// ---- 10_Core/90_Redundancy/FB_RedSync.TcPOU
FUNCTION_BLOCK FB_RedSync		// 동기화: 이 PLC의 운영 설정(GVL_PERSIST, 모듈 설정 묶음 제외)과 제어 모드 요청(PCS마다)을 EAP로 매 스캔 상대에게 보내고, 상대가 Active이고 내가 Active가 아닐 때 받은 값으로 내 설정을 맞춘다
(* - 보내는 값은 EAP 변수 1개: 운영 설정(_stTx, ST_RedSyncCfg). 받는 값도 같은 모양(_stRx)
   - 모듈 설정 묶음(GVL_PERSIST.g_stModuleSet)은 동기화하지 않음: HMI가 두 PLC 모두에 씀 (PLC가 꺼져 있던 동안 바꾼 값은 복귀 전에 HMI에서 다시 쓸 것)
   - 맞추기: i_bApply일 때만, 값이 다른 것만 덮어씀 (같으면 안 씀: 저장을 불필요하게 만들지 않음). 바꾼 것이 없으면 q_bInSync
   - 살아 있음: _stRx.nSeq가 i_tTimeout 안에 바뀌어야 함 (q_bFresh)
   - I/O(AT %I*·%Q)는 설치할 때 XAE에서 연결. 인스턴스는 RedundancyTask의 PRG_Redundancy에 둠. 두 PLC 프로그램이 같아야 함 *)
VAR_INPUT
	i_bUse			: BOOL;
	i_bApply		: BOOL;				// 받은 값을 내 설정에 덮어써도 됨 (내가 Active가 아니고 상대가 Active이며 통신 정상)
	i_tTimeout		: TIME := T#2S;		// 새 값이 이 시간 안에 안 오면 낡은 것
END_VAR
VAR_OUTPUT
	q_bInSync		: BOOL;				// 받은 값이 낡지 않았고 내 설정이 그와 같음 (i_bApply일 때만 TRUE)
	q_bFresh		: BOOL;				// 상대가 보낸 값이 낡지 않음
	q_nApplied		: UDINT;			// 받은 값으로 덮어쓴 횟수 (필드 단위)
END_VAR
VAR
	(* I/O: XAE에서 연결 *)
	_stTx			AT %Q* : ST_RedSyncCfg;
	_stRx			AT %I* : ST_RedSyncCfg;

	_nLastSeq		: UDINT;
	_tonFresh		: TON;
END_VAR
VAR_TEMP
	bNew			: BOOL;
	bEq				: BOOL;
END_VAR

IF NOT i_bUse THEN
	RETURN;
END_IF

(* 1) 보내기 *)
_stTx.nProtoVer	:= 1;
_stTx.nSeq		:= _stTx.nSeq + 1;
_stTx.nModeReq1	:= GVL_SITE.g_fbCtrlMode1.i_nModeReq;
_stTx.aeOpMode := GVL_PERSIST.g_aeOpMode;
_stTx.astGroupSet := GVL_PERSIST.g_astGroupSet;
_stTx.astManualPolicy := GVL_PERSIST.g_astManualPolicy;
_stTx.astSourceReg := GVL_PERSIST.g_astSourceReg;
_stTx.astLimitReg := GVL_PERSIST.g_astLimitReg;
_stTx.astPermitReg := GVL_PERSIST.g_astPermitReg;
_stTx.astCompReg := GVL_PERSIST.g_astCompReg;
_stTx.astRuleCfg := GVL_PERSIST.g_astRuleCfg;
_stTx.astOutputCfg := GVL_PERSIST.g_astOutputCfg;
_stTx.astUnitRuleReg := GVL_PERSIST.g_astUnitRuleReg;
_stTx.astBatRuleReg := GVL_PERSIST.g_astBatRuleReg;
_stTx.stCmdFilter := GVL_PERSIST.g_stCmdFilter;
_stTx.stManualCmdSet := GVL_PERSIST.g_stManualCmdSet;
_stTx.stSeqSet := GVL_PERSIST.g_stSeqSet;
_stTx.stBrokerWatch := GVL_PERSIST.g_stBrokerWatch;	// [9번 수정 2026-11-09: 추가]

(* 2) 받기: 새 값이 오는지 *)
bNew := _stRx.nSeq <> _nLastSeq;
_nLastSeq := _stRx.nSeq;
_tonFresh(IN := NOT bNew, PT := i_tTimeout);
q_bFresh := _stRx.nProtoVer = 1 AND _stRx.nSeq <> 0 AND NOT _tonFresh.Q;

(* 3) 맞추기: 내가 Active가 아니고 상대가 Active일 때만 다른 것만 덮어씀 *)
q_bInSync := FALSE;
IF i_bApply AND q_bFresh THEN
	bEq := TRUE;
	IF GVL_SITE.g_fbCtrlMode1.i_nModeReq <> _stRx.nModeReq1 THEN
		GVL_SITE.g_fbCtrlMode1.i_nModeReq := _stRx.nModeReq1;
		q_nApplied := q_nApplied + 1;
		bEq := FALSE;
	END_IF
	IF MEMCMP(ADR(GVL_PERSIST.g_aeOpMode), ADR(_stRx.aeOpMode), SIZEOF(_stRx.aeOpMode)) <> 0 THEN
		GVL_PERSIST.g_aeOpMode := _stRx.aeOpMode;
		q_nApplied := q_nApplied + 1;
		bEq := FALSE;
	END_IF
	IF MEMCMP(ADR(GVL_PERSIST.g_astGroupSet), ADR(_stRx.astGroupSet), SIZEOF(_stRx.astGroupSet)) <> 0 THEN
		GVL_PERSIST.g_astGroupSet := _stRx.astGroupSet;
		q_nApplied := q_nApplied + 1;
		bEq := FALSE;
	END_IF
	IF MEMCMP(ADR(GVL_PERSIST.g_astManualPolicy), ADR(_stRx.astManualPolicy), SIZEOF(_stRx.astManualPolicy)) <> 0 THEN
		GVL_PERSIST.g_astManualPolicy := _stRx.astManualPolicy;
		q_nApplied := q_nApplied + 1;
		bEq := FALSE;
	END_IF
	IF MEMCMP(ADR(GVL_PERSIST.g_astSourceReg), ADR(_stRx.astSourceReg), SIZEOF(_stRx.astSourceReg)) <> 0 THEN
		GVL_PERSIST.g_astSourceReg := _stRx.astSourceReg;
		q_nApplied := q_nApplied + 1;
		bEq := FALSE;
	END_IF
	IF MEMCMP(ADR(GVL_PERSIST.g_astLimitReg), ADR(_stRx.astLimitReg), SIZEOF(_stRx.astLimitReg)) <> 0 THEN
		GVL_PERSIST.g_astLimitReg := _stRx.astLimitReg;
		q_nApplied := q_nApplied + 1;
		bEq := FALSE;
	END_IF
	IF MEMCMP(ADR(GVL_PERSIST.g_astPermitReg), ADR(_stRx.astPermitReg), SIZEOF(_stRx.astPermitReg)) <> 0 THEN
		GVL_PERSIST.g_astPermitReg := _stRx.astPermitReg;
		q_nApplied := q_nApplied + 1;
		bEq := FALSE;
	END_IF
	IF MEMCMP(ADR(GVL_PERSIST.g_astCompReg), ADR(_stRx.astCompReg), SIZEOF(_stRx.astCompReg)) <> 0 THEN
		GVL_PERSIST.g_astCompReg := _stRx.astCompReg;
		q_nApplied := q_nApplied + 1;
		bEq := FALSE;
	END_IF
	IF MEMCMP(ADR(GVL_PERSIST.g_astRuleCfg), ADR(_stRx.astRuleCfg), SIZEOF(_stRx.astRuleCfg)) <> 0 THEN
		GVL_PERSIST.g_astRuleCfg := _stRx.astRuleCfg;
		q_nApplied := q_nApplied + 1;
		bEq := FALSE;
	END_IF
	IF MEMCMP(ADR(GVL_PERSIST.g_astOutputCfg), ADR(_stRx.astOutputCfg), SIZEOF(_stRx.astOutputCfg)) <> 0 THEN
		GVL_PERSIST.g_astOutputCfg := _stRx.astOutputCfg;
		q_nApplied := q_nApplied + 1;
		bEq := FALSE;
	END_IF
	IF MEMCMP(ADR(GVL_PERSIST.g_astUnitRuleReg), ADR(_stRx.astUnitRuleReg), SIZEOF(_stRx.astUnitRuleReg)) <> 0 THEN
		GVL_PERSIST.g_astUnitRuleReg := _stRx.astUnitRuleReg;
		q_nApplied := q_nApplied + 1;
		bEq := FALSE;
	END_IF
	IF MEMCMP(ADR(GVL_PERSIST.g_astBatRuleReg), ADR(_stRx.astBatRuleReg), SIZEOF(_stRx.astBatRuleReg)) <> 0 THEN
		GVL_PERSIST.g_astBatRuleReg := _stRx.astBatRuleReg;
		q_nApplied := q_nApplied + 1;
		bEq := FALSE;
	END_IF
	IF MEMCMP(ADR(GVL_PERSIST.g_stCmdFilter), ADR(_stRx.stCmdFilter), SIZEOF(_stRx.stCmdFilter)) <> 0 THEN
		GVL_PERSIST.g_stCmdFilter := _stRx.stCmdFilter;
		q_nApplied := q_nApplied + 1;
		bEq := FALSE;
	END_IF
	IF MEMCMP(ADR(GVL_PERSIST.g_stManualCmdSet), ADR(_stRx.stManualCmdSet), SIZEOF(_stRx.stManualCmdSet)) <> 0 THEN
		GVL_PERSIST.g_stManualCmdSet := _stRx.stManualCmdSet;
		q_nApplied := q_nApplied + 1;
		bEq := FALSE;
	END_IF
	IF MEMCMP(ADR(GVL_PERSIST.g_stSeqSet), ADR(_stRx.stSeqSet), SIZEOF(_stRx.stSeqSet)) <> 0 THEN
		GVL_PERSIST.g_stSeqSet := _stRx.stSeqSet;
		q_nApplied := q_nApplied + 1;
		bEq := FALSE;
	END_IF
	IF MEMCMP(ADR(GVL_PERSIST.g_stBrokerWatch), ADR(_stRx.stBrokerWatch), SIZEOF(_stRx.stBrokerWatch)) <> 0 THEN	// [9번 수정 2026-11-09: 추가]
		GVL_PERSIST.g_stBrokerWatch := _stRx.stBrokerWatch;
		q_nApplied := q_nApplied + 1;
		bEq := FALSE;
	END_IF
	q_bInSync := bEq;
END_IF

END_FUNCTION_BLOCK

// ---- 10_Core/90_Redundancy/FB_RedState.TcPOU
FUNCTION_BLOCK FB_RedState		// 이중화 상태 기계 (순수 로직). 역할 + 상대 상태 → 이 PLC가 Active인지, 장비에 써도 되는지. 두 PLC가 동시에 Active가 되지 않게 함
(* 규칙
   - 이중화를 안 쓰면 항상 Active이고 바로 쓴다
   - 역할 설정 오류(NoMatch) 또는 두 PLC 역할이 같음 → Failed (둘 다 장비에 쓰지 않음)
   - Primary: 시작하면 상대 상태를 볼 때까지 Init. 상대가 Active가 아니면 Active, 이미 Active이면 뺏지 않고 Standby
   - 절체: Secondary는 상대가 Lost(EAP·접점 둘 다 끊김)이고 tTakeoverDelay가 지나면 Active (Standby → Active)
   - 복귀: Primary가 Standby에서 상대(Secondary)가 Active이고 통신이 tFailbackStable 동안 정상이면 Handover(넘겨받기 요청)로 감.
     Secondary는 상대가 Handover이면 Active를 내려놓고 Standby로. Primary는 상대가 Active가 아니게 되면 Active.
     tHandoverTimeout 안에 안 내려놓으면 Primary가 Standby로 돌아가 다시 기다림. 둘 다 안 쓰는 틈이 생기지만 둘 다 쓰는 일은 없음
   - 둘 다 Active로 보이면 Secondary가 Standby로 물러남 (Primary 우선)
   - 상대 Active = EAP 하트비트의 Active (EAP 정상일 때) 또는 Active 접점 (접점 정상일 때)
   - PLC가 멈췄다 이어지면(i_bReset) Init부터 다시 정함: 멈춘 사이 상대가 Active를 넘겨받았을 수 있으므로 옛 Active를 이어 쓰지 않고, 상대 상태를 본 뒤 Standby로 들어가 복귀 절차를 밟음
   - 장비에 쓰는 허가(q_bWrite)는 Active가 된 뒤 tWriteHold가 지나야 켜짐 (승격 직후 계산이 안정되기를 기다림). Active가 아니게 되면 바로 꺼짐 *)
VAR_INPUT
	i_bUse			: BOOL;				// GVL_SITE.RED_SET.bUse
	i_stSet			: ST_RedSet;		// 시간 설정
	i_eRole			: E_RedRole;
	i_ePeer			: E_RedPeer;
	i_bPeerActive	: BOOL;				// 상대가 Active (EAP 또는 접점. 정상인 쪽만 반영해서 넘길 것)
	i_bPeerHandover	: BOOL;				// 상대가 Handover라고 알림 (EAP 정상일 때만)
	i_bRoleConflict	: BOOL;				// 두 PLC 역할이 같음 (FB_RedPeerMonitor)
	i_bReset		: BOOL;				// PLC가 멈췄다 이어짐: 상태를 Init부터 다시 정함 (멈춘 사이 상대가 Active를 넘겨받았을 수 있음)
	i_bSyncDone		: BOOL := TRUE;		// 복귀 전에 상대에게서 받을 값 동기화가 끝났음 (4단계에서 연결. 지금은 항상 TRUE)
END_VAR
VAR_OUTPUT
	q_eState		: E_RedState;
	q_bActive		: BOOL;				// Active 상태 (상대에게 알림)
	q_bWrite		: BOOL;				// 장비에 써도 됨 (Active + 쓰기 대기 지남)
	q_nSwitchCount	: UDINT;			// Active가 바뀐 횟수 (들어가거나 나옴)
	q_eLastSwitch	: E_RedSwitch;		// 마지막으로 바뀐 이유
END_VAR
VAR
	_ePrev			: E_RedState;
	_tonTakeover	: TON;
	_tonFailback	: TON;
	_tonHandover	: TON;
	_tonHold		: TON;
END_VAR

// 타이머는 매 스캔 부름
_tonTakeover(IN := i_eRole = E_RedRole.Secondary AND q_eState = E_RedState.Standby AND i_ePeer = E_RedPeer.Lost, PT := i_stSet.tTakeoverDelay);
_tonFailback(IN := i_eRole = E_RedRole.Primary AND q_eState = E_RedState.Standby AND i_ePeer = E_RedPeer.Alive AND i_bPeerActive AND i_bSyncDone, PT := i_stSet.tFailbackStable);
_tonHandover(IN := q_eState = E_RedState.Handover, PT := i_stSet.tHandoverTimeout);

IF i_bReset THEN
	q_eState := E_RedState.Init;
ELSIF NOT i_bUse THEN
	q_eState := E_RedState.Active;
ELSIF i_eRole = E_RedRole.NoMatch OR i_bRoleConflict THEN
	q_eState := E_RedState.Failed;
ELSIF i_eRole = E_RedRole.Reading THEN
	q_eState := E_RedState.Init;
ELSE
	IF q_eState = E_RedState.Failed THEN
		q_eState := E_RedState.Init;		// 오류가 풀리면 처음부터 다시 정함
	END_IF
	CASE q_eState OF
	E_RedState.Init:
		IF i_eRole = E_RedRole.Secondary THEN
			q_eState := E_RedState.Standby;
		ELSIF i_ePeer <> E_RedPeer.Unknown THEN		// Primary: 상대 상태를 본 뒤 정함
			IF i_bPeerActive THEN
				q_eState := E_RedState.Standby;
			ELSE
				q_eState := E_RedState.Active;
				q_eLastSwitch := E_RedSwitch.Start;
			END_IF
		END_IF
	E_RedState.Standby:
		IF i_eRole = E_RedRole.Secondary THEN
			IF _tonTakeover.Q THEN
				q_eState := E_RedState.Active;		// 절체
				q_eLastSwitch := E_RedSwitch.PeerLost;
			END_IF
		ELSIF i_ePeer <> E_RedPeer.Unknown THEN		// Primary
			IF NOT i_bPeerActive THEN
				q_eState := E_RedState.Active;		// 상대가 Active가 아님 (정지·대기)
				q_eLastSwitch := E_RedSwitch.Start;
			ELSIF _tonFailback.Q THEN
				q_eState := E_RedState.Handover;	// 복귀: 상대에게 Active를 내려놓으라고 알림
			END_IF
		END_IF
	E_RedState.Handover:
		IF NOT i_bPeerActive THEN
			q_eState := E_RedState.Active;			// 상대가 내려놓음 (또는 사라짐)
			q_eLastSwitch := E_RedSwitch.Failback;
		ELSIF _tonHandover.Q OR i_ePeer <> E_RedPeer.Alive THEN
			q_eState := E_RedState.Standby;			// 포기하고 처음부터 다시 기다림
		END_IF
	E_RedState.Active:
		IF i_eRole = E_RedRole.Secondary AND (i_bPeerActive OR i_bPeerHandover) THEN
			q_eState := E_RedState.Standby;			// Primary에 양보
			q_eLastSwitch := E_RedSwitch.Yield;
		END_IF
	ELSE
		q_eState := E_RedState.Init;
	END_CASE
END_IF

// Active가 들어가거나 나올 때 횟수
IF (q_eState = E_RedState.Active) <> (_ePrev = E_RedState.Active) THEN
	q_nSwitchCount := q_nSwitchCount + 1;
END_IF
_ePrev := q_eState;

q_bActive := q_eState = E_RedState.Active;
_tonHold(IN := q_bActive, PT := i_stSet.tWriteHold);
q_bWrite := q_bActive AND (_tonHold.Q OR NOT i_bUse);

END_FUNCTION_BLOCK

// ---- 10_Core/90_Redundancy/FB_RedLink.TcPOU
FUNCTION_BLOCK FB_RedLink		// 이중화 연결: EAP 하트비트 보내기·받기 + 접점 신호(EL2004 출력·EL1004 입력) 보내기·받기 + 상대 상태 판정 (FB_RedPeerMonitor)
(* - I/O 연결(AT %I*·%Q)은 설치할 때 XAE에서 한다. 인스턴스는 RedundancyTask를 도는 PRG_Redundancy에 둔다
   - EAP 보내기 _stTx → 상대가 받음, 받기 _stRx ← 상대가 보냄, Quality _nEapQuality: EAP 변수 연결 (값 = 마지막 갱신 뒤 지난 시간, 100 us 단위)
   - 접점: _bDoAlive(EL2004 채널 1)는 주기적으로 뒤집음 → 상대 _bDiPeerAlive(EL1004 채널 1). _bDoActive(채널 2)는 이 PLC가 Active인 동안 TRUE → 상대 _bDiPeerActive(채널 2)
   - 두 PLC에 같은 프로그램을 넣고, 두 PLC의 I/O 연결이 서로 마주 보게 한다 *)
VAR_INPUT
	i_stSet			: ST_RedSet;
	i_eRole			: E_RedRole;
	i_bActive		: BOOL;
	i_eState		: E_RedState;		// 이 PLC의 이중화 상태 (상대에게 알림)
END_VAR
VAR_OUTPUT
	q_ePeer			: E_RedPeer;		// 상대 상태
	q_bEapOk		: BOOL;
	q_bWireOk		: BOOL;
	q_stPeer		: ST_RedHeartbeat;	// 상대가 보낸 역할·Active (EAP 정상일 때만)
	q_bPeerWireActive: BOOL;			// 상대 Active 접점 (EAP와 따로 보는 값)
	q_bRoleConflict	: BOOL;				// 두 PLC 역할이 같음
	q_nTxCount		: UDINT;			// 보낸 하트비트 수
END_VAR
VAR CONSTANT
	PULSE_HALF		: TIME := T#100MS;	// alive 접점을 뒤집는 간격 (접점 타임아웃보다 충분히 짧게)
END_VAR
VAR
	(* I/O: XAE에서 연결 *)
	_stTx			AT %Q* : ST_RedHeartbeat;
	_stRx			AT %I* : ST_RedHeartbeat;
	_nEapQuality	AT %I* : UINT;		// EAP Subscriber의 Quality = 갱신 안 된 시간 (100 us 단위). tEapTimeout 이하면 정상
	_bDoAlive		AT %Q* : BOOL;		// EL2004 채널 1
	_bDoActive		AT %Q* : BOOL;		// EL2004 채널 2
	_bDiPeerAlive	AT %I* : BOOL;		// EL1004 채널 1
	_bDiPeerActive	AT %I* : BOOL;		// EL1004 채널 2

	_fbMon			: FB_RedPeerMonitor;
	_tonPulse		: TON;
END_VAR

(* 1) 보내기 *)
q_nTxCount			:= q_nTxCount + 1;
_stTx.nProtoVer		:= 2;
_stTx.nCounter		:= q_nTxCount;
_stTx.nRole			:= TO_INT(i_eRole);
_stTx.bActive		:= i_bActive;
_stTx.nState		:= TO_INT(i_eState);

_tonPulse(IN := NOT _tonPulse.Q, PT := PULSE_HALF);		// Q가 한 스캔 켜질 때마다 뒤집음
IF _tonPulse.Q THEN
	_bDoAlive := NOT _bDoAlive;
END_IF
_bDoActive			:= i_bActive;

(* 2) 받아서 판정 *)
_fbMon(	i_stRx			:= _stRx,
		i_nMyRole		:= TO_INT(i_eRole),
		i_bEapQualityOk	:= UINT_TO_UDINT(_nEapQuality) <= TIME_TO_UDINT(i_stSet.tEapTimeout) * 10,	// Quality = 갱신 안 된 시간 (100 us 단위)
		i_bWireAlive	:= _bDiPeerAlive,
		i_tEapTimeout	:= i_stSet.tEapTimeout,
		i_tWireTimeout	:= i_stSet.tWireTimeout,
		i_tStartGrace	:= i_stSet.tStartGrace);
q_ePeer				:= _fbMon.q_ePeer;
q_bEapOk			:= _fbMon.q_bEapOk;
q_bWireOk			:= _fbMon.q_bWireOk;
q_stPeer			:= _fbMon.q_stPeer;
q_bPeerWireActive	:= _bDiPeerActive;
q_bRoleConflict		:= _fbMon.q_bRoleConflict;

END_FUNCTION_BLOCK

// ---- 10_Core/90_Redundancy/FB_RedPeerMonitor.TcPOU
FUNCTION_BLOCK FB_RedPeerMonitor		// 상대 PLC 상태 판정 (순수 로직: I/O를 직접 안 봄). EAP 하트비트(카운터가 바뀌고 Quality 정상)와 접점 신호(값이 바뀜)를 따로 보고 합침
// 판정 규칙: 둘 다 정상 = Alive, 한쪽만 끊김 = 그 통신 고장 (상대는 살아 있음, 절체 안 함), 둘 다 끊김 = Lost (절체 조건)
VAR_INPUT
	i_stRx			: ST_RedHeartbeat;	// 받은 EAP 하트비트
	i_bEapQualityOk	: BOOL;				// EAP Quality가 정상
	i_nMyRole		: INT;				// 이 PLC의 역할 (E_RedRole). 받은 역할이 같으면 내 프레임이 되돌아온 것으로 보고 무시
	i_bWireAlive	: BOOL;				// 상대 alive 접점(DI)의 지금 값. 상대가 주기적으로 뒤집음
	i_tEapTimeout	: TIME := T#500MS;	// 카운터가 이 시간 안 바뀌면 EAP 끊김
	i_tWireTimeout	: TIME := T#500MS;	// 접점이 이 시간 안 바뀌면 접점 끊김
	i_tStartGrace	: TIME := T#3S;		// 시작 직후 대기: 이 안에는 아직 못 봐도 Unknown
END_VAR
VAR_OUTPUT
	q_ePeer			: E_RedPeer;
	q_bEapOk		: BOOL;				// EAP 하트비트 정상
	q_bWireOk		: BOOL;				// 접점 신호 정상
	q_stPeer		: ST_RedHeartbeat;	// 상대가 보낸 값. EAP가 정상일 때만 채움 (아니면 0)
	q_bRoleConflict	: BOOL;				// 상대가 나와 같은 역할로 살아 있음 (두 PLC 역할 설정 오류). 접점도 살아 있을 때만 (내 프레임이 되돌아온 경우와 구분)
END_VAR
VAR
	_bInit			: BOOL;
	_nLastCount		: UDINT;
	_bLastWire		: BOOL;
	_bEapSeen		: BOOL;			// 시작 뒤 카운터가 바뀌는 것을 한 번이라도 봄
	_bWireSeen		: BOOL;
	_bSameSeen		: BOOL;
	_tonSame		: TON;
	_tonEap			: TON;
	_tonWire		: TON;
	_tonStart		: TON;
END_VAR
VAR_TEMP
	bEapMoved		: BOOL;
	bFromSelf		: BOOL;
	bSameMoved		: BOOL;
	bCntMoved		: BOOL;
	bWireMoved		: BOOL;
	stZero			: ST_RedHeartbeat;
END_VAR

IF NOT _bInit THEN
	_nLastCount	:= i_stRx.nCounter;
	_bLastWire	:= i_bWireAlive;
	_bInit		:= TRUE;
END_IF

// EAP: 카운터가 바뀌었고 Quality 정상이면 살아 있음. 안 바뀌는 시간이 길면 끊김 (상대 PLC가 멈추면 마지막 값이 그대로 남으므로 Quality만으로는 못 잡음)
bFromSelf		:= i_stRx.nRole = i_nMyRole;	// 상대와 내 역할은 항상 다름. 같으면 루프로 되돌아온 내 프레임 (또는 역할 설정 오류)
bCntMoved		:= i_bEapQualityOk AND i_stRx.nCounter <> _nLastCount;
bEapMoved		:= bCntMoved AND NOT bFromSelf;
_nLastCount		:= i_stRx.nCounter;
IF bEapMoved THEN
	_bEapSeen := TRUE;
END_IF
// 같은 역할 프레임이 계속 오는지 (Primary·Secondary일 때만. 시작 중 Reading끼리는 제외)
bSameMoved		:= bCntMoved AND bFromSelf AND (i_nMyRole = 1 OR i_nMyRole = 2);
IF bSameMoved THEN
	_bSameSeen := TRUE;
END_IF
_tonSame(IN := NOT bSameMoved, PT := i_tEapTimeout);
_tonEap(IN := NOT bEapMoved, PT := i_tEapTimeout);
q_bEapOk		:= _bEapSeen AND NOT _tonEap.Q AND i_bEapQualityOk AND NOT bFromSelf;

// 접점: 값이 바뀌면 살아 있음
bWireMoved		:= i_bWireAlive <> _bLastWire;
_bLastWire		:= i_bWireAlive;
IF bWireMoved THEN
	_bWireSeen := TRUE;
END_IF
_tonWire(IN := NOT bWireMoved, PT := i_tWireTimeout);
q_bWireOk		:= _bWireSeen AND NOT _tonWire.Q;
q_bRoleConflict	:= _bSameSeen AND NOT _tonSame.Q AND q_bWireOk;

_tonStart(IN := TRUE, PT := i_tStartGrace);

IF q_bEapOk AND q_bWireOk THEN
	q_ePeer := E_RedPeer.Alive;
ELSIF q_bWireOk THEN
	q_ePeer := E_RedPeer.EapLost;
ELSIF q_bEapOk THEN
	q_ePeer := E_RedPeer.WireLost;
ELSIF NOT _bEapSeen AND NOT _bWireSeen AND NOT _tonStart.Q THEN
	q_ePeer := E_RedPeer.Unknown;
ELSE
	q_ePeer := E_RedPeer.Lost;
END_IF

IF q_bEapOk THEN
	q_stPeer := i_stRx;
ELSE
	q_stPeer := stZero;
END_IF

END_FUNCTION_BLOCK

// ---- 20_Module/Common/FB_AuxIo.TcPOU
FUNCTION_BLOCK FB_AuxIo EXTENDS FB_DeviceBase IMPLEMENTS I_AuxDevice		// 벡호프 단자 I/O (EL1xxx 입력, EL2xxx 출력, EL3xxx 아날로그 입력, EL4xxx 아날로그 출력)
(* 점은 TwinCAT 화면에서 _abDi·_abDo·_anAi·_anAo 칸에 하나씩 연결. 점 번호 = 배열 칸 번호
   이 FB를 PlcTask가 아닌 태스크에서 쓰면 그 태스크 PRG 안에 선언 (GVL에 두면 TcContextName 필요) *)
VAR_INPUT
	i_afAiGain		: ARRAY[1..GVL_PARAM.AUX_AI_MAX] OF REAL;		// 아날로그 입력 = 원시값 × 배율 + 오프셋. 배율 0 = 1 (예: PT100 EL3202는 0.1)
	i_afAiOffset	: ARRAY[1..GVL_PARAM.AUX_AI_MAX] OF REAL;
	i_afAoGain		: ARRAY[1..GVL_PARAM.AUX_AO_MAX] OF REAL;		// 아날로그 출력 원시값 = 값 / 배율. 배율 0 = 1
END_VAR
VAR
	_abDi	AT %I*	: ARRAY[1..GVL_PARAM.AUX_DI_MAX] OF BOOL;
	_abDo	AT %Q*	: ARRAY[1..GVL_PARAM.AUX_DO_MAX] OF BOOL;
	_anAi	AT %I*	: ARRAY[1..GVL_PARAM.AUX_AI_MAX] OF INT;
	_anAo	AT %Q*	: ARRAY[1..GVL_PARAM.AUX_AO_MAX] OF INT;
	_bWcError AT %I* : BOOL;		// (선택) EtherCAT WcState 연결. 안 연결하면 늘 정상
END_VAR

METHOD M_Cycle
IF NOT _bWcError THEN
	M_MarkAlive();
END_IF
M_UpdateComm();
END_METHOD

PROPERTY Comm : BOOL
GET
Comm := _bComm;
END_GET
END_PROPERTY

METHOD M_GetBit : BOOL
VAR_INPUT
	i_nPoint	: UINT;
END_VAR
IF i_nPoint >= 1 AND i_nPoint <= GVL_PARAM.AUX_DI_MAX THEN
	M_GetBit := _abDi[i_nPoint];
END_IF
END_METHOD

METHOD M_GetValue : ST_Val
VAR_INPUT
	i_nPoint	: UINT;
END_VAR
IF i_nPoint >= 1 AND i_nPoint <= GVL_PARAM.AUX_AI_MAX THEN
	M_GetValue.fValue := INT_TO_REAL(_anAi[i_nPoint]) * SEL(i_afAiGain[i_nPoint] = 0, i_afAiGain[i_nPoint], 1.0) + i_afAiOffset[i_nPoint];
	M_GetValue.bValid := _bComm;
END_IF
END_METHOD

METHOD M_SetBit
VAR_INPUT
	i_nPoint	: UINT;
	i_bValue	: BOOL;
END_VAR
IF i_nPoint >= 1 AND i_nPoint <= GVL_PARAM.AUX_DO_MAX THEN
	_abDo[i_nPoint] := i_bValue;
END_IF
END_METHOD

METHOD M_SetValue
VAR_INPUT
	i_nPoint	: UINT;
	i_fValue	: REAL;
END_VAR
IF i_nPoint >= 1 AND i_nPoint <= GVL_PARAM.AUX_AO_MAX THEN
	// [결함 13 수정 2026-11-04: 값·게인이 숫자가 아니면 0 (LIMIT·REAL_TO_INT에서 FPU 예외). 원래 아래 줄만]
	IF F_RealOk(i_fValue) AND F_RealOk(i_afAoGain[i_nPoint]) THEN
		_anAo[i_nPoint] := REAL_TO_INT(LIMIT(-32768.0, i_fValue / SEL(i_afAoGain[i_nPoint] = 0, i_afAoGain[i_nPoint], 1.0), 32767.0));
	ELSE
		_anAo[i_nPoint] := 0;
	END_IF
END_IF
END_METHOD

END_FUNCTION_BLOCK

// ---- 10_Core/03_Base/FB_DeviceBase.TcPOU
FUNCTION_BLOCK ABSTRACT FB_DeviceBase EXTENDS FB_ModuleBase
VAR_INPUT
	i_tCommTimeout		: TIME := T#10S;	// 이 시간 동안 정상 응답이 없으면 통신 이상
	i_tReadPeriod		: TIME := T#200MS;	// 읽기 주기. 장비마다 GVL_SITE 인스턴스 선언에서 바꿈 (i_tCommTimeout보다 짧게)
END_VAR
VAR
	_bComm				: BOOL;		// 통신 정상
	_bAlive				: BOOL;		// 이번 스캔에 정상 응답(또는 하트비트 변화)이 있었음
	_bEverAlive			: BOOL;		// 부팅 후 한 번이라도 응답이 있었음
	_tonCommLoss		: TON;
	_fbRead				: FB_ReadTimer;
	_nWriteFails		: UINT;		// 잇달아 실패한 쓰기 수
	_bWriteFail			: BOOL;		// 쓰기 실패 (드라이버가 상태 bWriteFail에 넣음)
END_VAR
VAR CONSTANT
	WRITE_FAIL_COUNT	: UINT := 3;	// 쓰기가 이만큼 잇달아 실패하면 쓰기 실패로 봄 (한 번 성공하면 풀림)
END_VAR

METHOD PROTECTED M_MarkAlive
_bAlive		:= TRUE;
_bEverAlive	:= TRUE;
END_METHOD

METHOD PROTECTED M_IsReadTime : BOOL		// 읽을 때가 되면 TRUE (i_tReadPeriod마다). 스캔당 한 번만 부를 것
_fbRead(i_tPeriod := i_tReadPeriod);
M_IsReadTime := _fbRead.q_bDue;
END_METHOD

METHOD PROTECTED M_UpdateComm
// 마지막 정상 응답 이후 i_tCommTimeout이 지나면 통신 이상
_tonCommLoss(IN := NOT _bAlive, PT := i_tCommTimeout);
_bComm	:= _bEverAlive AND NOT _tonCommLoss.Q;	// 한 번도 응답이 없으면 정상으로 보지 않는다
_bAlive	:= FALSE;								// 다음 스캔을 위해 초기화
END_METHOD

METHOD PROTECTED M_MarkWriteResult		// 쓰기 결과를 알림 (드라이버가 쓰기 응답을 받을 때마다). 잇달아 WRITE_FAIL_COUNT번 실패하면 _bWriteFail, 한 번 성공하면 풀림
VAR_INPUT
	i_bOk	: BOOL;
END_VAR
IF i_bOk THEN
	_nWriteFails	:= 0;
	_bWriteFail		:= FALSE;
ELSE
	IF _nWriteFails < WRITE_FAIL_COUNT THEN
		_nWriteFails := _nWriteFails + 1;
	END_IF
	_bWriteFail := _nWriteFails >= WRITE_FAIL_COUNT;
END_IF
END_METHOD

END_FUNCTION_BLOCK

// ---- 10_Core/02_Util/FB_ReadTimer.TcPOU
FUNCTION_BLOCK FB_ReadTimer		// 읽기 주기 타이머: 읽을 때가 되면 그 스캔만 q_bDue = TRUE. 처음 호출 때 바로 TRUE
VAR_INPUT
	i_tPeriod		: TIME := T#200MS;	// 읽기 주기. T#0S면 매 스캔
END_VAR
VAR_OUTPUT
	q_bDue			: BOOL;
END_VAR
VAR
	_bStarted		: BOOL;
	_tonWait		: TON;
END_VAR

// 스캔당 한 번만 호출할 것
_tonWait(IN := _bStarted, PT := i_tPeriod);
q_bDue := NOT _bStarted OR _tonWait.Q;

IF q_bDue THEN
	_bStarted := TRUE;
	_tonWait(IN := FALSE, PT := i_tPeriod);	// 이번 스캔부터 다시 셈
	_tonWait(IN := TRUE, PT := i_tPeriod);
END_IF

END_FUNCTION_BLOCK

// ---- 20_Module/Mqtt/FB_SrcEms.TcPOU
FUNCTION_BLOCK FB_SrcEms EXTENDS FB_SourceBase		// 지령원: EMS (상위 플랫폼, MQTT command). 명령 핸들러(FB_EmsCommand)가 해석한 명령을 요청으로 냄
(* - 입력 i_stCmd는 MAIN(A_PassEmsCmd)이 GVL_IF에서 일관되게 복사해 넘긴다. 이 FB는 GVL을 보지 않는다
   - 상태 명령(PCS Run·Standby·Stop·EStop·Reset, 배터리 Close·Open): 번호가 바뀌면 새 명령. 큐에 넣고 스캔마다 1개씩 요청으로 낸다.
     받는 운전 모드는 등록표 stStateMode가 정한다. 배터리 Reset은 운전자 리셋(PCS Reset, 전체)으로 낸다
   - 충전·방전 P 지령: PCS 한 대의 kW를 그 PCS의 유닛들에 정격 비율로 나눠 유닛 지령(astUnit)으로 낸다.
     i_bPEnable이 TRUE일 때만 낸다 (기본 FALSE). 제어 모드(FB_CtrlModeMgr)와 어떻게 묶을지는 정해지면 여기서 연결 (상태 명령은 이 값과 무관하게 받음)
   - 새 메시지(nRxCount)나 새 명령이 만료 시간(등록 tExpire) 안에 오면 살아 있음. 끊기면 P 지령·요청 큐를 버린다 (돌아와도 옛 지령이 되살아나지 않음)
   - PMS가 켜진 뒤 처음 복사본은 번호만 맞춘다 (재기동 때 지난 명령을 실행하지 않음)
   - 배터리 비상정지(EStop)는 지령원 요청 종류에 없어 받지 않고 q_nUnsupported로 센다 *)
VAR_INPUT
	i_stCmd			: ST_IfEmsCmd;	// MAIN이 GVL_IF에서 복사한 명령 칸
	i_bValid		: BOOL;			// i_stCmd가 한 번이라도 일관되게 복사됨
	i_astUnitCfg	: ARRAY[1..GVL_PARAM.UNIT_COUNT] OF ST_UnitCfg;	// 유닛 ← PCS 번호 (명령은 PCS 번호로 옴)
	i_astBmsCfg		: ARRAY[1..GVL_PARAM.BMS_COUNT] OF ST_BmsCfg;	// BMS → 배터리 그룹
	i_bPEnable		: BOOL;			// 충전·방전 P 지령을 낼지 (기본 FALSE. 제어 모드와의 연결 방식이 정해질 때까지 끔)
END_VAR
VAR_OUTPUT
	q_nUnsupported	: UDINT;		// 받을 수 없는 명령 수 (배터리 비상정지)
	q_nQueueDrop	: UDINT;		// 큐가 가득 차 버린 요청 수
END_VAR
VAR CONSTANT
	QUEUE_PCS		: UINT := 16;
	QUEUE_BAT		: UINT := 8;
END_VAR
VAR
	_bSynced		: BOOL;
	_nRxCount		: UDINT;
	_anPcsSeq		: ARRAY[1..GVL_PARAM.PCS_COUNT] OF UDINT;
	_anPSeq			: ARRAY[1..GVL_PARAM.PCS_COUNT] OF UDINT;
	_anBatSeq		: ARRAY[1..GVL_PARAM.BMS_COUNT] OF UDINT;
	_abUnitP		: ARRAY[1..GVL_PARAM.UNIT_COUNT] OF BOOL;	// 이 유닛에 받아 둔 P 지령 있음
	_afUnitP		: ARRAY[1..GVL_PARAM.UNIT_COUNT] OF REAL;	// kW, 유닛 출력 (방전 +)
	_astPcsQ		: ARRAY[1..QUEUE_PCS] OF ST_PcsReq;
	_nPcsHead		: UINT := 1;
	_nPcsCount		: UINT;
	_astBatQ		: ARRAY[1..QUEUE_BAT] OF ST_BatReq;
	_nBatHead		: UINT := 1;
	_nBatCount		: UINT;
END_VAR

METHOD PRIVATE M_PushBat
VAR_INPUT
	i_eCmd		: E_BatCmd;
	i_nBatGroup	: UINT;
END_VAR
VAR
	nTail		: UINT;
END_VAR
IF _nBatCount >= QUEUE_BAT THEN
	q_nQueueDrop := q_nQueueDrop + 1;
	RETURN;
END_IF
nTail := ((_nBatHead + _nBatCount - 1) MOD QUEUE_BAT) + 1;
_astBatQ[nTail].eCmd		:= i_eCmd;
_astBatQ[nTail].nBatGroup	:= i_nBatGroup;
_nBatCount := _nBatCount + 1;
END_METHOD

METHOD PRIVATE M_PushPcs
VAR_INPUT
	i_eCmd		: E_PcsCmd;
	i_nUnit		: UINT;		// 0 = 그룹 전체
END_VAR
VAR
	nTail		: UINT;
END_VAR
IF _nPcsCount >= QUEUE_PCS THEN
	q_nQueueDrop := q_nQueueDrop + 1;
	RETURN;
END_IF
nTail := ((_nPcsHead + _nPcsCount - 1) MOD QUEUE_PCS) + 1;
_astPcsQ[nTail].eCmd	:= i_eCmd;
_astPcsQ[nTail].nUnit	:= i_nUnit;
_nPcsCount := _nPcsCount + 1;
END_METHOD

METHOD M_ReasonText : WSTRING(63)
VAR_INPUT
	i_nReason	: UINT;
END_VAR
M_ReasonText := "EMS 지령";
END_METHOD

METHOD M_UpdateOutput : BOOL
VAR
	p			: UINT;
	u			: UINT;
	b			: UINT;
	bFresh		: BOOL;
	bNewP		: BOOL;
	bAlgoOn		: BOOL;
	fSum		: REAL;
END_VAR
M_UpdateOutput := FALSE;

// 복사본이 아직 한 번도 없으면 기다림. 처음 받은 복사본은 번호만 맞춤 (지난 명령을 실행하지 않음)
IF NOT i_bValid THEN
	RETURN;
END_IF
IF NOT _bSynced THEN
	_bSynced := TRUE;
	_nRxCount := i_stCmd.nRxCount;
	FOR p := 1 TO GVL_PARAM.PCS_COUNT DO
		_anPcsSeq[p]	:= i_stCmd.astPcs[p].nSeq;
		_anPSeq[p]		:= i_stCmd.anPcsPSeq[p];
	END_FOR
	FOR b := 1 TO GVL_PARAM.BMS_COUNT DO
		_anBatSeq[b]	:= i_stCmd.astBat[b].nSeq;
	END_FOR
	RETURN;
END_IF

// 끊긴 상태(지난 스캔 기준)면 받아 둔 P 지령과 큐를 버림
IF _tonExpire.Q THEN
	FOR u := 1 TO GVL_PARAM.UNIT_COUNT DO
		_abUnitP[u] := FALSE;
	END_FOR
	_nPcsCount := 0;
	_nBatCount := 0;
END_IF

bFresh := FALSE;
bNewP := FALSE;
IF i_stCmd.nRxCount <> _nRxCount THEN
	_nRxCount := i_stCmd.nRxCount;
	bFresh := TRUE;
END_IF

// PCS: 상태 명령 → 그 PCS의 유닛마다 요청 (리셋은 전체 한 번), P 지령 → 유닛에 정격 비율로 나눔
FOR p := 1 TO GVL_PARAM.PCS_COUNT DO
	IF i_stCmd.astPcs[p].nSeq <> _anPcsSeq[p] THEN
		_anPcsSeq[p] := i_stCmd.astPcs[p].nSeq;
		bFresh := TRUE;
		IF i_stCmd.astPcs[p].eCmd = E_PcsCmd.Reset THEN
			M_PushPcs(E_PcsCmd.Reset, 0);
		ELSIF i_stCmd.astPcs[p].eCmd <> E_PcsCmd.None THEN
			FOR u := 1 TO GVL_PARAM.UNIT_COUNT DO
				IF i_astUnitCfg[u].nPcs = p THEN
					M_PushPcs(i_stCmd.astPcs[p].eCmd, u);
				END_IF
			END_FOR
		END_IF
	END_IF
	IF i_stCmd.anPcsPSeq[p] <> _anPSeq[p] THEN
		_anPSeq[p] := i_stCmd.anPcsPSeq[p];
		bFresh := TRUE;
		bNewP := TRUE;
		fSum := 0.0;
		FOR u := 1 TO GVL_PARAM.UNIT_COUNT DO
			IF i_astUnitCfg[u].nPcs = p THEN
				fSum := fSum + i_astUnitCfg[u].fPRated;
			END_IF
		END_FOR
		FOR u := 1 TO GVL_PARAM.UNIT_COUNT DO
			IF i_astUnitCfg[u].nPcs = p THEN
				_abUnitP[u] := TRUE;
				IF fSum > 0.0 THEN
					_afUnitP[u] := i_stCmd.afPcsP[p] * i_astUnitCfg[u].fPRated / fSum;
				ELSE
					_afUnitP[u] := 0.0;
				END_IF
			END_IF
		END_FOR
	END_IF
END_FOR

// BMS: 투입·개방은 배터리 그룹 요청, 리셋은 운전자 리셋
FOR b := 1 TO GVL_PARAM.BMS_COUNT DO
	IF i_stCmd.astBat[b].nSeq <> _anBatSeq[b] THEN
		_anBatSeq[b] := i_stCmd.astBat[b].nSeq;
		bFresh := TRUE;
		IF i_stCmd.astBat[b].eCmd = E_BatCmd.Close OR i_stCmd.astBat[b].eCmd = E_BatCmd.Open THEN
			M_PushBat(i_stCmd.astBat[b].eCmd, i_astBmsCfg[b].nBatGroup);
		ELSIF i_stCmd.astBat[b].eCmd = E_BatCmd.Reset THEN
			M_PushPcs(E_PcsCmd.Reset, 0);
		ELSE
			q_nUnsupported := q_nUnsupported + 1;
		END_IF
	END_IF
END_FOR

// 큐에서 한 스캔에 하나씩 요청으로 냄
IF _nPcsCount > 0 THEN
	_stOut.stPcsReq := _astPcsQ[_nPcsHead];
	_nPcsHead := (_nPcsHead MOD QUEUE_PCS) + 1;
	_nPcsCount := _nPcsCount - 1;
END_IF
IF _nBatCount > 0 THEN
	_stOut.stBatReq := _astBatQ[_nBatHead];
	_nBatHead := (_nBatHead MOD QUEUE_BAT) + 1;
	_nBatCount := _nBatCount - 1;
END_IF

// P 지령: 알고리즘이 선택된 그룹에서만. 받은 값은 새 명령이 올 때까지 유지 (만료되면 위에서 버림)
bAlgoOn := i_bPEnable;		// 등록 사용 여부(bEnable)는 FB_SourceBase가 처리 (꺼져 있으면 전부 지움)
FOR u := 1 TO GVL_PARAM.UNIT_COUNT DO
	_stOut.astUnit[u].bPSetActive	:= _abUnitP[u] AND bAlgoOn;
	_stOut.astUnit[u].fPSet			:= _afUnitP[u];
	_stOut.astUnit[u].bQSetActive	:= FALSE;
END_FOR
_stOut.bNewSet := bNewP AND bAlgoOn;

M_UpdateOutput := bFresh;
END_METHOD

END_FUNCTION_BLOCK

// ---- 20_Module/Driver/Plaspo/FB_PlaspoPcs.TcPOU
FUNCTION_BLOCK FB_PlaspoPcs EXTENDS FB_DeviceBase IMPLEMENTS I_Pcs		// 플라스포 PCS (Modbus TCP, 유닛 1개). 레지스터 맵은 Helios FB_PlaspoPcs와 같음
(* ---------------------------------------------------------------
   상태 (읽기 맵 → ST_UnitState)
   - 고장 비트 → Fault, 인버터 정지 → Stop
   - 운전 중이면서 마지막 상태 명령이 Standby → Standby, 그 밖의 운전 중 → Run
     (플라스포에는 Standby 상태가 따로 없어서 "운전 중 + 대기 모드(103 = 0)"를 Standby로 봄)
   명령 (레지스터: 값)
   - 기동    101: 55, 105: 1       - 정지·비상정지 101: 99, 105: 1 (비상정지 명령이 따로 없음)
   - 리셋    102: 33, 105: 1       - Standby  (정지 중이면 기동 먼저) 106: 1, 103: 0, 107: 0
   - 출력    P > 0 방전 103: 2, P < 0 충전 103: 1, 107: |P| × i_fPScale. 방향이 같으면 107만 씀
   - Q 지령은 이 맵에 없음 → 무시
   쓰기: 한 번에 레지스터 하나, 사이 간격 i_tWriteGap. 상태 명령이 출력보다 먼저.
         출력은 가장 최근 값만 보냄 (밀려 있으면 덮어씀)
   현장 확인: 유효전력 부호(i_bPInvert), 출력 레지스터 단위(i_fPScale)
   --------------------------------------------------------------- *)
VAR_INPUT
	i_sIpAddr		: STRING(15);
	i_nPort			: UINT := 502;
	i_nUnitId		: BYTE := 1;
	i_fPScale		: REAL := 1.0;		// 출력 레지스터(107) = kW × 배율
	i_bPInvert		: BOOL := TRUE;		// 읽은 유효전력 부호 뒤집기 (Helios: -acActive → 방전 +)
	i_tWriteGap		: TIME := T#300MS;	// 레지스터 쓰기 사이 간격 (Helios 300 ms)
	i_tTimeout		: TIME := T#1S;
END_VAR
VAR
	(* 읽기 *)
	_fbMbRead			: FB_MBReadRegs;
	_stReadMap			: ST_PlaspoPcsRaw;
	_bReadDue		: BOOL;
	_bReading		: BOOL;
	_bReadError		: BOOL;
	_nReadErrId		: UDINT;
	_stUnit			: ST_UnitState;
	_bStandbyMode	: BOOL;				// 마지막 상태 명령이 Standby
	(* 보낼 목록 (대기): 상태 명령은 가장 최근 것만, 출력은 가장 최근 값만 *)
	_anCmdRegAddr		: ARRAY[1..5] OF UINT;	// 보낼 상태 명령 (가장 최근 것만)
	_anCmdRegValue		: ARRAY[1..5] OF INT;
	_nCmdRegCount		: UINT;				// 0 = 없음
	_bPowerPending	: BOOL;
	_nPowerDir		: INT;				// 보낼 방향 (103 값): 0 그대로, 1 충전, 2 방전
	_nPowerAbs	: INT;				// 107
	_nDirWritten	: INT;				// 마지막으로 쓴 103
	(* 지금 보내는 목록 *)
	_fbMbWrite		: FB_MBWriteRegs;
	_anSendAddr		: ARRAY[1..5] OF UINT;
	_anSendValue		: ARRAY[1..5] OF INT;
	_nSendCount		: UINT;
	_nSendIdx		: UINT;
	_nWriteStep		: UINT;				// 0 다음 일 고르기, 1 쓰기 시작, 2 끝나기 기다림, 3 간격
	_bWriteError	: BOOL;
	_nWriteErrId	: UDINT;
	_tonWriteGap			: TON;
	_nCopyIdx			: UINT;				// 액션에서 쓰는 반복 변수
END_VAR

ACTION A_MapToUnitState:
_stUnit.bComm		:= _bComm AND NOT _stReadMap.nPcsStatus.5;
_stUnit.bFault		:= _stReadMap.nPcsStatus.1;
_stUnit.bCtrlReady	:= _stReadMap.nRemoteMode = 1;

IF NOT _stUnit.bComm THEN
	_stUnit.eRunState := E_RunState.Unknown;
ELSIF _stUnit.bFault THEN
	_stUnit.eRunState := E_RunState.Fault;
ELSIF NOT _stReadMap.nPcsStatus.0 THEN
	_stUnit.eRunState := E_RunState.Stop;
ELSIF _bStandbyMode THEN
	_stUnit.eRunState := E_RunState.Standby;
ELSE
	_stUnit.eRunState := E_RunState.Run;
END_IF

_stUnit.stP.fValue	:= INT_TO_REAL(_stReadMap.nAcActive) * 0.1 * SEL(i_bPInvert, 1.0, -1.0);
_stUnit.stP.bValid	:= _stUnit.bComm;
_stUnit.stQ.fValue	:= INT_TO_REAL(_stReadMap.nAcReactive) * 0.1;
_stUnit.stQ.bValid	:= _stUnit.bComm;
END_ACTION

ACTION A_ReadRegisters:
// 읽기 주기마다 한 번 (Helios A_ReadPcsData와 같은 순서)
IF NOT _bReading THEN
	IF _bReadDue THEN
		_fbMbRead(sIPAddr := i_sIpAddr, nTCPPort := i_nPort, nUnitID := i_nUnitId,
				nQuantity := SIZEOF(_stReadMap) / 2, nMBAddr := 1, cbLength := SIZEOF(_stReadMap),
				pDestAddr := ADR(_stReadMap), tTimeout := i_tTimeout, bExecute := TRUE);
		_bReading := TRUE;
	END_IF
ELSE
	_fbMbRead(bExecute := FALSE);
	IF NOT _fbMbRead.bBusy THEN
		_bReadError	:= _fbMbRead.bError;
		_nReadErrId	:= _fbMbRead.nErrId;
		IF NOT _fbMbRead.bError THEN
			M_MarkAlive();
		END_IF
		_bReading := FALSE;
	END_IF
END_IF
END_ACTION

ACTION A_WriteQueue:
CASE _nWriteStep OF
	0:	// 다음 일: 상태 명령이 먼저, 그다음 출력
		_nSendCount := 0;
		IF _nCmdRegCount > 0 THEN
			FOR _nCopyIdx := 1 TO _nCmdRegCount DO
				_anSendAddr[_nCopyIdx]	:= _anCmdRegAddr[_nCopyIdx];
				_anSendValue[_nCopyIdx]	:= _anCmdRegValue[_nCopyIdx];
			END_FOR
			_nSendCount := _nCmdRegCount;
			_nCmdRegCount := 0;
		ELSIF _bPowerPending THEN
			IF _nPowerDir <> 0 AND _nPowerDir <> _nDirWritten THEN
				_anSendAddr[1] := 106;	_anSendValue[1] := 1;
				_anSendAddr[2] := 103;	_anSendValue[2] := _nPowerDir;
				_anSendAddr[3] := 107;	_anSendValue[3] := _nPowerAbs;
				_nSendCount := 3;
			ELSE
				_anSendAddr[1] := 107;	_anSendValue[1] := _nPowerAbs;
				_nSendCount := 1;
			END_IF
			_bPowerPending := FALSE;
		END_IF
		IF _nSendCount > 0 THEN
			_nSendIdx	:= 1;
			_nWriteStep	:= 1;
		END_IF

	1:	// 레지스터 하나 쓰기 시작
		_fbMbWrite(sIPAddr := i_sIpAddr, nTCPPort := i_nPort, nUnitID := i_nUnitId,
				 nQuantity := 1, nMBAddr := _anSendAddr[_nSendIdx], cbLength := 2,
				 pSrcAddr := ADR(_anSendValue[_nSendIdx]), tTimeout := i_tTimeout, bExecute := TRUE);
		_nWriteStep := 2;

	2:	// 끝나기 기다림
		_fbMbWrite(bExecute := FALSE);
		IF NOT _fbMbWrite.bBusy THEN
			_bWriteError := _fbMbWrite.bError;
			_nWriteErrId := _fbMbWrite.nErrId;
			IF NOT _fbMbWrite.bError AND _anSendAddr[_nSendIdx] = 103 THEN
				_nDirWritten := _anSendValue[_nSendIdx];
			END_IF
			IF _fbMbWrite.bError THEN
				_nSendIdx := _nSendCount;		// 실패하면 이 일은 그만 (상태 명령은 시퀀서가 다시 보냄)
			END_IF
			_nWriteStep := 3;
		END_IF

	3:	// 간격
		_tonWriteGap(IN := TRUE, PT := i_tWriteGap);
		IF _tonWriteGap.Q THEN
			_tonWriteGap(IN := FALSE);
			IF _nSendIdx < _nSendCount THEN
				_nSendIdx	:= _nSendIdx + 1;
				_nWriteStep	:= 1;
			ELSE
				_nWriteStep	:= 0;
			END_IF
		END_IF
END_CASE
END_ACTION

METHOD M_Cycle
_bReadDue := M_IsReadTime();
A_ReadRegisters();
M_UpdateComm();
A_MapToUnitState();
A_WriteQueue();
END_METHOD

METHOD M_GetUnitState : ST_UnitState
VAR_INPUT
	i_nSub		: UINT;
END_VAR
IF i_nSub = 1 THEN
	M_GetUnitState := _stUnit;
END_IF
END_METHOD

METHOD PRIVATE M_QueueCmdAndApply		// 상태 명령 보낼 목록을 새로 만듦: 명령 레지스터 하나 + 적용 신호(105 ← 1)
VAR_INPUT
	i_nAddr		: UINT;
	i_nValue	: INT;
END_VAR
_nCmdRegCount := 0;
M_QueueRegister(i_nAddr, i_nValue);
M_QueueRegister(105, 1);
END_METHOD

METHOD PRIVATE M_QueueRegister		// 상태 명령 보낼 목록에 레지스터 하나(주소 ← 값) 추가
VAR_INPUT
	i_nAddr		: UINT;
	i_nValue	: INT;
END_VAR
IF _nCmdRegCount < 5 THEN
	_nCmdRegCount := _nCmdRegCount + 1;
	_anCmdRegAddr[_nCmdRegCount]	:= i_nAddr;
	_anCmdRegValue[_nCmdRegCount]	:= i_nValue;
END_IF
END_METHOD

METHOD M_SetPower : BOOL
VAR_INPUT
	i_nSub		: UINT;
	i_fP		: REAL;			// kW, 방전 +
	i_fQ		: REAL;			// 이 맵에는 Q 지령이 없음
END_VAR
IF i_nSub <> 1 THEN
	RETURN;
END_IF
IF i_fP > 0.05 THEN
	_nPowerDir := 2;			// 방전
ELSIF i_fP < -0.05 THEN
	_nPowerDir := 1;			// 충전
ELSE
	_nPowerDir := 0;			// 0 kW: 방향은 그대로 두고 107만
END_IF
// [결함 13 수정 2026-11-04: 지령·배율이 숫자가 아니면 0 (LIMIT·REAL_TO_INT에서 FPU 예외). 원래 _nPowerAbs := REAL_TO_INT(LIMIT(0.0, ABS(i_fP) * i_fPScale, 32767.0));]
IF F_RealOk(i_fP) AND F_RealOk(i_fPScale) THEN
	_nPowerAbs	:= REAL_TO_INT(LIMIT(0.0, ABS(i_fP) * i_fPScale, 32767.0));
ELSE
	_nPowerAbs	:= 0;
END_IF
_bPowerPending	:= TRUE;
M_SetPower := TRUE;
END_METHOD

METHOD M_SetStateCmd : BOOL
VAR_INPUT
	i_nSub		: UINT;
	i_stCmd		: ST_PcsCmd;
END_VAR
IF i_nSub <> 1 THEN
	RETURN;
END_IF

CASE i_stCmd.eCmd OF
	E_PcsCmd.Run:
		_bStandbyMode := FALSE;
		_nDirWritten := 0;			// 첫 출력 때 방향(103)을 다시 씀
		IF _stUnit.eRunState = E_RunState.Stop THEN
			M_QueueCmdAndApply(101, 55);			// 기동
		END_IF
		// 이미 운전 중이면 쓸 것 없음: Run으로 보고하고 출력 지령을 따름

	E_PcsCmd.Standby:
		_bStandbyMode := TRUE;
		_nCmdRegCount := 0;
		IF _stUnit.eRunState = E_RunState.Stop THEN
			M_QueueRegister(101, 55);
			M_QueueRegister(105, 1);
		END_IF
		M_QueueRegister(106, 1);
		M_QueueRegister(103, 0);
		M_QueueRegister(107, 0);

	E_PcsCmd.Stop,
	E_PcsCmd.EStop:
		_bStandbyMode := FALSE;
		_nDirWritten := 0;
		M_QueueCmdAndApply(101, 99);

	E_PcsCmd.Reset:
		M_QueueCmdAndApply(102, 33);
ELSE
	RETURN;
END_CASE
M_SetStateCmd := TRUE;
END_METHOD

PROPERTY RawMap : ST_PlaspoPcsRaw		// 마지막으로 읽은 레지스터 맵 (보고 매핑용. 제어에 쓰지 않음)
GET
RawMap := _stReadMap;
END_GET
END_PROPERTY

END_FUNCTION_BLOCK

// ---- 20_Module/Virtual/FB_PcsSim.TcPOU
FUNCTION_BLOCK FB_PcsSim EXTENDS FB_DeviceBase IMPLEMENTS I_Pcs		// 가상 PCS (시험용)
VAR_INPUT
	i_tTau			: TIME := T#500MS;	// 출력 응답 시정수
	i_bForceFault	: BOOL;				// 시험: 전 유닛 고장
	i_bForceLocal	: BOOL;				// 시험: 로컬 모드 (PMS 제어 불가)
	i_bForceCommLoss	: BOOL;			// 시험: 통신 끊김 (응답 안 함. i_tCommTimeout 뒤 통신 이상)
	i_bIgnoreCmd	: BOOL;				// 시험: 상태 명령을 접수하되 상태는 바꾸지 않음 (P/Q 지령은 적용)
	i_bFaultFlagOnly	: BOOL;			// 시험: 운전 상태는 그대로 두고 고장 표시만 켬 (해제도 이 입력으로 함)
END_VAR
VAR
	_aeState		: ARRAY[1..GVL_PARAM.MAX_SUB] OF E_RunState;
	_afPSet			: ARRAY[1..GVL_PARAM.MAX_SUB] OF REAL;
	_afQSet			: ARRAY[1..GVL_PARAM.MAX_SUB] OF REAL;
	_afbPLag			: ARRAY[1..GVL_PARAM.MAX_SUB] OF FB_Lpf;
	_afbQLag			: ARRAY[1..GVL_PARAM.MAX_SUB] OF FB_Lpf;
	_astUnit		: ARRAY[1..GVL_PARAM.MAX_SUB] OF ST_UnitState;
END_VAR

METHOD M_Cycle
VAR
	u		: UINT;
	fPTarget		: REAL;
	fQTarget		: REAL;
END_VAR
IF M_IsReadTime() AND NOT i_bForceCommLoss THEN		// 읽기 주기마다 응답한 것으로 봄 (시험: 통신 끊김이면 응답 안 함)
	M_MarkAlive();
END_IF
M_UpdateComm();

FOR u := 1 TO GVL_PARAM.MAX_SUB DO
	IF _aeState[u] = E_RunState.Unknown THEN
		_aeState[u] := E_RunState.Stop;
	END_IF
	IF i_bForceFault THEN
		_aeState[u] := E_RunState.Fault;
	END_IF

	// 운전 중이면 지령을, 아니면 0을 1차 지연으로 따라감
	IF _aeState[u] = E_RunState.Run THEN
		fPTarget := _afPSet[u];
		fQTarget := _afQSet[u];
	ELSE
		fPTarget := 0;
		fQTarget := 0;
	END_IF
	_afbPLag[u](i_fIn := fPTarget, i_tTau := i_tTau);
	_afbQLag[u](i_fIn := fQTarget, i_tTau := i_tTau);

	_astUnit[u].bComm		:= _bComm;
	_astUnit[u].eRunState	:= _aeState[u];
	_astUnit[u].bCtrlReady	:= NOT i_bForceLocal;
	_astUnit[u].bFault		:= (_aeState[u] = E_RunState.Fault) OR i_bFaultFlagOnly;
	_astUnit[u].stP.fValue	:= _afbPLag[u].q_fOut;
	_astUnit[u].stP.bValid	:= TRUE;
	_astUnit[u].stQ.fValue	:= _afbQLag[u].q_fOut;
	_astUnit[u].stQ.bValid	:= TRUE;
END_FOR
END_METHOD

METHOD M_GetUnitState : ST_UnitState
VAR_INPUT
	i_nSub		: UINT;
END_VAR
IF i_nSub >= 1 AND i_nSub <= GVL_PARAM.MAX_SUB THEN
	M_GetUnitState := _astUnit[i_nSub];
END_IF
END_METHOD

METHOD M_SetPower : BOOL
VAR_INPUT
	i_nSub		: UINT;
	i_fP		: REAL;
	i_fQ		: REAL;
END_VAR
IF i_nSub < 1 OR i_nSub > GVL_PARAM.MAX_SUB THEN
	RETURN;
END_IF
_afPSet[i_nSub] := i_fP;
_afQSet[i_nSub] := i_fQ;
M_SetPower := TRUE;
END_METHOD

METHOD M_SetStateCmd : BOOL
VAR_INPUT
	i_nSub		: UINT;
	i_stCmd		: ST_PcsCmd;
END_VAR
IF i_nSub < 1 OR i_nSub > GVL_PARAM.MAX_SUB THEN
	RETURN;
END_IF

CASE i_stCmd.eCmd OF
	E_PcsCmd.Run:
		IF NOT i_bIgnoreCmd AND _aeState[i_nSub] <> E_RunState.Fault THEN _aeState[i_nSub] := E_RunState.Run; END_IF

	E_PcsCmd.Standby:
		IF NOT i_bIgnoreCmd AND _aeState[i_nSub] <> E_RunState.Fault THEN _aeState[i_nSub] := E_RunState.Standby; END_IF

	E_PcsCmd.Stop,
	E_PcsCmd.EStop:
		IF NOT i_bIgnoreCmd AND _aeState[i_nSub] <> E_RunState.Fault THEN _aeState[i_nSub] := E_RunState.Stop; END_IF

	E_PcsCmd.Reset:
		IF NOT i_bIgnoreCmd AND _aeState[i_nSub] = E_RunState.Fault AND NOT i_bForceFault THEN _aeState[i_nSub] := E_RunState.Stop; END_IF
ELSE
	RETURN;		// 배터리 명령 등은 PCS가 받지 않음
END_CASE

M_SetStateCmd := TRUE;
END_METHOD

END_FUNCTION_BLOCK

// ---- 20_Module/Report/FB_RptPlaspoPcs.TcPOU
FUNCTION_BLOCK FB_RptPlaspoPcs		// 보고 매핑: 플라스포 PCS 읽기값 + 코어 결과 → MQTT pcs 발행 레코드 (보고 전용, 제어에 쓰지 않음)
(* 필드 대응 (플라스포 읽기 맵 ST_PlaspoPcsRaw, 괄호는 레지스터 번호):
   SystemOperationMode  코어 운전 모드 (Manual 0, Auto 1)
   OperationMode        nOpMode (4) 그대로
   PMSActivePower       PMS가 이 PCS에 낸 지령 kW (분배 결과. 장비 쓰기를 막아도 나옴)
   RemoteMode           nRemoteMode (3)
   Status               nPcsStatus (1) 그대로: bit0 운전, bit1 고장, bit2 경고, bit5 PCS 내부 통신 이상
   AcActivePower·AcReactivePower  드라이버가 변환한 P·Q (방전 +, 0.1 kW·kvar)
   PowerFactor          nAcPf (29) × i_fPfScale
   Frequency            nAcFreq (26) × 0.1
   AcRs·St·TrVoltage    anAcVolt[1..3] (20~22) × i_fVoltScale  (선간 전압으로 가정)
   AcR·S·TVoltage       읽지 않음 → 0
   AcR·S·TCurrent       anAcCurrent[1..3] (23~25) × i_fCurrScale
   DcLinkVoltage·DcVoltage  nDcLinkVolt (36)·nDcVolt (37) × i_fDcVoltScale
   DcCurrent            nDcCurrent (38) × i_fDcCurrScale
   DcActivePower        nDcPower (39) × i_fDcPowerScale
   InsulationResistance 읽지 않음 → 0
   Temperature1~4       anIgbtTemp[1..4] (12~15) × i_fTempScale
   Temperature5~8       anAcFilterTemp[1..4] (16~19) × i_fTempScale
   Warning1             anFault[5] (11). Warning2~10 → 0
   Fault1~4             anFault[1..4] (7~10). Fault5~10 → 0
   통신이 끊기면 레코드 전체가 0 (이 값만으로는 끊김을 알 수 없으니 GVL_IF.g_stReport.abPcsComm을 봄)
   배율(i_f…Scale)은 레지스터 맵 문서로 확인되지 않은 값이라 기본 1.0 (= 레지스터 값 그대로). 실제 값과 비교해 맞출 것 *)
VAR_INPUT
	i_stRaw			: ST_PlaspoPcsRaw;	// 드라이버 FB_PlaspoPcs.RawMap
	i_stUnit		: ST_UnitState;		// 이 PCS의 유닛 상태 (FB_Snapshot)
	i_eOpMode		: E_OpMode;			// 이 유닛의 실제 운전 모드 (FB_ModeSwitch)
	i_fPCmd			: REAL;				// kW, PMS가 낸 지령 (FB_Distributor 유닛 지령)
	i_fPfScale		: REAL := 1.0;
	i_fVoltScale	: REAL := 1.0;
	i_fCurrScale	: REAL := 1.0;
	i_fDcVoltScale	: REAL := 1.0;
	i_fDcCurrScale	: REAL := 1.0;
	i_fDcPowerScale	: REAL := 1.0;
	i_fTempScale	: REAL := 1.0;
END_VAR
VAR_OUTPUT
	q_stPcs			: ST_PcsPublish_V1;	// 발행 직전 레코드 (DeviceIndex는 PRG_Mqtt가 채움)
	q_bComm			: BOOL;				// 통신 정상
END_VAR
VAR
	_stNone			: ST_PcsPublish_V1;
END_VAR

q_stPcs := _stNone;
q_bComm := i_stUnit.bComm;
IF NOT q_bComm THEN
	RETURN;
END_IF

IF i_eOpMode = E_OpMode.Auto THEN
	q_stPcs.SystemOperationMode := 1;
ELSE
	q_stPcs.SystemOperationMode := 0;
END_IF
q_stPcs.OperationMode		:= UINT_TO_UDINT(i_stRaw.nOpMode);
q_stPcs.PMSActivePower		:= i_fPCmd;
q_stPcs.RemoteMode			:= UINT_TO_UDINT(i_stRaw.nRemoteMode);
q_stPcs.Status				:= DWORD_TO_UDINT(WORD_TO_DWORD(i_stRaw.nPcsStatus));

q_stPcs.AcActivePower		:= i_stUnit.stP.fValue;
q_stPcs.AcReactivePower		:= i_stUnit.stQ.fValue;
q_stPcs.PowerFactor			:= INT_TO_REAL(i_stRaw.nAcPf) * i_fPfScale;
q_stPcs.Frequency			:= UINT_TO_REAL(i_stRaw.nAcFreq) * 0.1;

q_stPcs.AcRsVoltage			:= UINT_TO_REAL(i_stRaw.anAcVolt[1]) * i_fVoltScale;
q_stPcs.AcStVoltage			:= UINT_TO_REAL(i_stRaw.anAcVolt[2]) * i_fVoltScale;
q_stPcs.AcTrVoltage			:= UINT_TO_REAL(i_stRaw.anAcVolt[3]) * i_fVoltScale;
q_stPcs.AcRCurrent			:= UINT_TO_REAL(i_stRaw.anAcCurrent[1]) * i_fCurrScale;
q_stPcs.AcSCurrent			:= UINT_TO_REAL(i_stRaw.anAcCurrent[2]) * i_fCurrScale;
q_stPcs.AcTCurrent			:= UINT_TO_REAL(i_stRaw.anAcCurrent[3]) * i_fCurrScale;

q_stPcs.DcLinkVoltage		:= UINT_TO_REAL(i_stRaw.nDcLinkVolt) * i_fDcVoltScale;
q_stPcs.DcVoltage			:= UINT_TO_REAL(i_stRaw.nDcVolt) * i_fDcVoltScale;
q_stPcs.DcCurrent			:= INT_TO_REAL(i_stRaw.nDcCurrent) * i_fDcCurrScale;
q_stPcs.DcActivePower		:= INT_TO_REAL(i_stRaw.nDcPower) * i_fDcPowerScale;

q_stPcs.Temperature1		:= INT_TO_REAL(i_stRaw.anIgbtTemp[1]) * i_fTempScale;
q_stPcs.Temperature2		:= INT_TO_REAL(i_stRaw.anIgbtTemp[2]) * i_fTempScale;
q_stPcs.Temperature3		:= INT_TO_REAL(i_stRaw.anIgbtTemp[3]) * i_fTempScale;
q_stPcs.Temperature4		:= INT_TO_REAL(i_stRaw.anIgbtTemp[4]) * i_fTempScale;
q_stPcs.Temperature5		:= INT_TO_REAL(i_stRaw.anAcFilterTemp[1]) * i_fTempScale;
q_stPcs.Temperature6		:= INT_TO_REAL(i_stRaw.anAcFilterTemp[2]) * i_fTempScale;
q_stPcs.Temperature7		:= INT_TO_REAL(i_stRaw.anAcFilterTemp[3]) * i_fTempScale;
q_stPcs.Temperature8		:= INT_TO_REAL(i_stRaw.anAcFilterTemp[4]) * i_fTempScale;

q_stPcs.Warning1			:= DWORD_TO_UDINT(WORD_TO_DWORD(i_stRaw.anFault[5]));
q_stPcs.Fault1				:= DWORD_TO_UDINT(WORD_TO_DWORD(i_stRaw.anFault[1]));
q_stPcs.Fault2				:= DWORD_TO_UDINT(WORD_TO_DWORD(i_stRaw.anFault[2]));
q_stPcs.Fault3				:= DWORD_TO_UDINT(WORD_TO_DWORD(i_stRaw.anFault[3]));
q_stPcs.Fault4				:= DWORD_TO_UDINT(WORD_TO_DWORD(i_stRaw.anFault[4]));

END_FUNCTION_BLOCK

// ---- 20_Module/Driver/Esolution/FB_EsolutionBms.TcPOU
FUNCTION_BLOCK FB_EsolutionBms EXTENDS FB_DeviceBase IMPLEMENTS I_Bms

VAR_INPUT
 i_bEnable : BOOL;
 i_sIpAddr : STRING(15);
 i_nPort : UINT := 502;
 i_nUnitId : BYTE := 1;
 i_tTimeout : TIME := T#1S;
 i_bWritePermit : BOOL; // site dispatcher: config OK AND active PLC
END_VAR
VAR_OUTPUT
 q_eRequestResult : E_UpsResult;
 q_nTransportError : UDINT;
END_VAR
VAR
 _fbJob : FB_UpsModbusJob;
 _bLaunch : BOOL;
 _bCurrentWrite : BOOL;
 _bDiscardResponse : BOOL; // response started before a disable must not complete a new snapshot
 _nFunction : UINT;
 _nAddress : WORD;
 _nQuantity : WORD;
 _wValue : WORD;
 _bPendingWrite : BOOL;
 _nPendingAddress : WORD;
 _wPendingValue : WORD;
 _nPendingQty : WORD; // 1 = FC06, 2~3 = FC16 같은 값 여러 칸 [2026-11-13]
 _awValues : ARRAY[0..2] OF WORD;
 _nPoll : UINT;
 _nCopy : UINT;
 _bReadDue : BOOL;
END_VAR

VAR_INPUT
 i_nRackCount : UINT := 1; // configure actual installed count, max10
 i_nModuleCount : UINT := GVL_PARAM.MODULES_PER_RACK; // installed modules; map stride remains 17 slots
 i_bReadDetails : BOOL := FALSE; // enable after unused module-slot response is confirmed
 i_tHeartbeatTimeout : TIME := T#10S;
 i_tDetailTimeout : TIME := T#60S;
END_VAR
VAR_OUTPUT
 q_stRaw : ST_EsolutionRaw;
 q_stState : ST_EsolutionState;
END_VAR
VAR
 _stWork : ST_EsolutionRaw;
 _stBat : ST_BatState;
 _nSampleSeq : UDINT;
 _nRack : UINT;
 _nOffset : UINT;
 _nDetailRack : UINT := 1;
 _nDetailOffset : UINT;
 _nDetailChunk : UINT;
 _wHeartbeat : WORD;
 _bHeartbeatChanged : BOOL;
 _tonHeartbeat : TON;
 _atonDetail : ARRAY[1..10] OF TON;
 _abDetailUpdated : ARRAY[1..10] OF BOOL;
 _wInstalledMask : WORD;
 _nLastRackCount : UINT;
 _nLastCoreCmdSeq : UDINT;
 _bHaveCoreCmd : BOOL;
END_VAR

METHOD M_Cycle
_bReadDue := M_IsReadTime();
IF NOT i_bEnable THEN
 _bDiscardResponse:=_bDiscardResponse OR _fbJob.q_bBusy;
 _bLaunch:=FALSE;
END_IF
IF NOT i_bEnable OR NOT i_bWritePermit OR NOT GVL_PARAM.UPS_CONTROL_ENABLED THEN
 _bPendingWrite := FALSE;
 // A queued but not yet started FC06 must not survive a gate transition.
 IF _bLaunch AND _bCurrentWrite THEN _bLaunch := FALSE; END_IF
END_IF
_fbJob(i_sIpAddr:=i_sIpAddr,i_nPort:=i_nPort,i_nUnitId:=i_nUnitId,i_tTimeout:=i_tTimeout,
 i_bExecute:=_bLaunch,i_bWritePermit:=i_bWritePermit AND i_bEnable,
 i_nFunction:=_nFunction,i_nAddress:=_nAddress,i_nQuantity:=_nQuantity,i_wValue:=_wValue,i_awValues:=_awValues);
_bLaunch := FALSE;
IF _fbJob.q_bDone THEN
 q_nTransportError := _fbJob.q_nErrorId;
 IF _bCurrentWrite THEN M_MarkWriteResult(NOT _fbJob.q_bError); END_IF
END_IF

IF i_nRackCount<1 OR i_nRackCount>10 OR i_nModuleCount<1 OR i_nModuleCount>17 THEN
 _bLaunch:=FALSE; _bPendingWrite:=FALSE;
 q_stState.bComm:=FALSE; q_stState.bValid:=FALSE; _stBat.bComm:=FALSE;
 RETURN;
END_IF
IF _nLastRackCount<>i_nRackCount THEN
 _nLastRackCount:=i_nRackCount; _nDetailRack:=1; _nDetailOffset:=0;
 FOR _nRack:=1 TO 10 DO q_stState.abDetailValid[_nRack]:=FALSE; END_FOR
END_IF
_bHeartbeatChanged:=FALSE;
FOR _nRack:=1 TO 10 DO _abDetailUpdated[_nRack]:=FALSE; END_FOR
IF _fbJob.q_bDone AND _bDiscardResponse THEN
 _bDiscardResponse:=FALSE; _nPoll:=0;
ELSIF _fbJob.q_bDone AND NOT _bCurrentWrite THEN
 IF _fbJob.q_bError THEN
  IF _nPoll=3 THEN _nDetailOffset:=0; END_IF
  _nPoll:=0;
 ELSE
  CASE _nPoll OF
   0: FOR _nCopy:=0 TO 26 DO _stWork.awSystem[_nCopy]:=_fbJob.q_awData[_nCopy]; END_FOR
   1: FOR _nCopy:=0 TO 39 DO _stWork.awRackAnalog[_nCopy]:=_fbJob.q_awData[_nCopy]; END_FOR
   2:
    FOR _nCopy:=0 TO 89 DO _stWork.awRackStatus[_nCopy]:=_fbJob.q_awData[_nCopy]; END_FOR
    q_stRaw.awSystem:=_stWork.awSystem;
    q_stRaw.awRackAnalog:=_stWork.awRackAnalog;
    q_stRaw.awRackStatus:=_stWork.awRackStatus;
    _bHeartbeatChanged:=_nSampleSeq=0 OR _wHeartbeat<>q_stRaw.awSystem[0];
    _wHeartbeat:=q_stRaw.awSystem[0]; _nSampleSeq:=F_UpsNextSeq(_nSampleSeq); M_MarkAlive();
   3:
    FOR _nCopy:=0 TO _nDetailChunk-1 DO
     _stWork.aawDetail[_nDetailRack,_nDetailOffset+_nCopy]:=_fbJob.q_awData[_nCopy];
    END_FOR
    IF _nDetailOffset+_nDetailChunk=406 THEN
     FOR _nCopy:=0 TO 405 DO q_stRaw.aawDetail[_nDetailRack,_nCopy]:=_stWork.aawDetail[_nDetailRack,_nCopy]; END_FOR
     q_stState.anDetailSeq[_nDetailRack]:=F_UpsNextSeq(q_stState.anDetailSeq[_nDetailRack]);
     _abDetailUpdated[_nDetailRack]:=TRUE;
     q_stState.abDetailValid[_nDetailRack]:=TRUE;
     _nDetailOffset:=0;
     IF _nDetailRack>=i_nRackCount THEN _nDetailRack:=1; ELSE _nDetailRack:=_nDetailRack+1; END_IF
    ELSE _nDetailOffset:=_nDetailOffset+_nDetailChunk; END_IF
  END_CASE
  IF _nPoll=3 OR (_nPoll=2 AND NOT i_bReadDetails) THEN _nPoll:=0; ELSE _nPoll:=_nPoll+1; END_IF
 END_IF
END_IF
M_UpdateComm();
_tonHeartbeat(IN:=NOT _bHeartbeatChanged,PT:=i_tHeartbeatTimeout);
// System Data 1~27
q_stState.nHeartbeat:=q_stRaw.awSystem[0]; // 1. 하트비트
q_stState.fVoltageV:=WORD_TO_REAL(q_stRaw.awSystem[1])*0.1; // 2. 전체 전압 (V)
q_stState.fCurrentA:=F_UpsSignedWord(q_stRaw.awSystem[2])*0.1; // 3. 전체 전류 (A)
q_stState.fSocPct:=WORD_TO_REAL(q_stRaw.awSystem[3])*0.1; // 4. 충전 상태 (%)
q_stState.fSohPct:=WORD_TO_REAL(q_stRaw.awSystem[4]); // 5. 건강 상태 (%)
q_stState.fChargePowerKw:=WORD_TO_REAL(q_stRaw.awSystem[5]); // 6. 충전 전력 (kW)
q_stState.fDischargePowerKw:=WORD_TO_REAL(q_stRaw.awSystem[6]); // 7. 방전 전력 (kW)
q_stState.fMaxCellVoltageMv:=WORD_TO_REAL(q_stRaw.awSystem[7]); // 8. 최대 셀 전압 (mV)
q_stState.fMinCellVoltageMv:=WORD_TO_REAL(q_stRaw.awSystem[8]); // 9. 최소 셀 전압 (mV)
q_stState.fAvgCellVoltageMv:=WORD_TO_REAL(q_stRaw.awSystem[9]); // 10. 평균 셀 전압 (mV)
q_stState.nMaxCellVoltageLocation:=q_stRaw.awSystem[10]; // 11. 최대 셀 전압 위치
q_stState.nMinCellVoltageLocation:=q_stRaw.awSystem[11]; // 12. 최소 셀 전압 위치
q_stState.fMaxCellTemperatureC:=F_UpsSignedWord(q_stRaw.awSystem[12])*0.1; // 13. 최고 셀 온도 (℃)
q_stState.fMinCellTemperatureC:=F_UpsSignedWord(q_stRaw.awSystem[13])*0.1; // 14. 최저 셀 온도 (℃)
q_stState.fAvgCellTemperatureC:=F_UpsSignedWord(q_stRaw.awSystem[14])*0.1; // 15. 평균 셀 온도 (℃)
q_stState.nMaxCellTemperatureLocation:=q_stRaw.awSystem[15]; // 16. 최고 셀 온도 위치
q_stState.nMinCellTemperatureLocation:=q_stRaw.awSystem[16]; // 17. 최저 셀 온도 위치
q_stState.fMaxRackSocPct:=WORD_TO_REAL(q_stRaw.awSystem[17])*0.1; // 18. 최대 랙 SOC (%)
q_stState.fMinRackSocPct:=WORD_TO_REAL(q_stRaw.awSystem[18])*0.1; // 19. 최소 랙 SOC (%)
q_stState.fMaxRackVoltageV:=WORD_TO_REAL(q_stRaw.awSystem[19])*0.1; // 20. 최대 랙 전압 (V)
q_stState.fMinRackVoltageV:=WORD_TO_REAL(q_stRaw.awSystem[20])*0.1; // 21. 최소 랙 전압 (V)
q_stState.fChargeLimitKw:=WORD_TO_REAL(q_stRaw.awSystem[21]); // 22. 충전 허용 전력 (kW)
q_stState.fDischargeLimitKw:=WORD_TO_REAL(q_stRaw.awSystem[22]); // 23. 방전 허용 전력 (kW)
q_stState.fChargeCurrentLimitA:=WORD_TO_REAL(q_stRaw.awSystem[23]); // 24. 충전 허용 전류 (A)
q_stState.fDischargeCurrentLimitA:=WORD_TO_REAL(q_stRaw.awSystem[24]); // 25. 방전 허용 전류 (A)
q_stState.wSystemContactor:=q_stRaw.awSystem[25]; // 26. 시스템 컨택터 상태 (맵 v1.4)
q_stState.wRackContactor:=q_stRaw.awSystem[26]; // 27. 랙 컨택터 상태 (맵 v1.4)
q_stState.bChargeContactorClosed:=q_stRaw.awSystem[25].0;
q_stState.bDischargeContactorClosed:=q_stRaw.awSystem[25].1;

q_stState.bComm:=_bComm AND i_bEnable;
q_stState.bFresh:=q_stState.bComm AND NOT _tonHeartbeat.Q;
q_stState.bValid:=q_stState.bFresh AND _nSampleSeq<>0;
q_stState.bWriteFail:=_bWriteFail;
q_stState.nSampleSeq:=_nSampleSeq;
q_stState.nRackCount:=i_nRackCount;
q_stState.nModuleCount:=i_nModuleCount;
q_stState.bWarn:=FALSE; q_stState.bFault:=FALSE; q_stState.bSystemLock:=FALSE;
FOR _nRack:=1 TO 10 DO
 _atonDetail[_nRack](IN:=NOT _abDetailUpdated[_nRack],PT:=i_tDetailTimeout);
 IF _atonDetail[_nRack].Q OR NOT q_stState.bValid OR NOT i_bReadDetails OR _nRack>i_nRackCount THEN
  q_stState.abDetailValid[_nRack]:=FALSE;
 END_IF
 IF _nRack<=i_nRackCount THEN
  _nOffset:=(_nRack-1)*9;
  q_stState.bWarn:=q_stState.bWarn OR (q_stRaw.awRackStatus[_nOffset] AND 16#01FF)<>0
   OR (q_stRaw.awRackStatus[_nOffset+2] AND 16#03FF)<>0 OR q_stRaw.awRackStatus[_nOffset+4].9;
  q_stState.bFault:=q_stState.bFault OR (q_stRaw.awRackStatus[_nOffset+3] AND 16#3FFF)<>0
   OR (q_stRaw.awRackStatus[_nOffset+4] AND 16#05FF)<>0 OR q_stRaw.awRackStatus[_nOffset+5]<>0
   OR (q_stRaw.awRackStatus[_nOffset+6] AND 16#00FF)<>0 OR (q_stRaw.awRackStatus[_nOffset+7] AND 16#8001)<>0;
  q_stState.bSystemLock:=q_stState.bSystemLock OR q_stRaw.awRackStatus[_nOffset].8 OR q_stRaw.awRackStatus[_nOffset+3].13;
 END_IF
END_FOR
// 컨택터 상태는 맵 v1.4 Input 26·27로 판단 (명령이나 운전 모드로 추정하지 않음) [2026-11-13]
// 붙음 = 설치 랙 중 하나라도 붙음 AND 충전·방전 중 하나라도 붙음 (배터리가 버스에 이어짐).
// 그래서 하나라도 붙어 있으면 코어 개방(Open)이 나가고, 개방 확인은 다 떨어져야 됨.
q_stState.bContactorFeedbackKnown:=q_stState.bValid;
_wInstalledMask:=SHL(WORD#1,i_nRackCount)-1;
_stBat.bComm:=q_stState.bValid;
_stBat.bContactorClosed:=q_stState.bValid AND (q_stState.wRackContactor AND _wInstalledMask)<>0
 AND (q_stState.bChargeContactorClosed OR q_stState.bDischargeContactorClosed);
_stBat.bWarn:=q_stState.bWarn; _stBat.bFault:=q_stState.bFault; _stBat.bSysStop:=q_stState.bSystemLock;
_stBat.stSoc.fValue:=q_stState.fSocPct;
_stBat.stSoc.bValid:=q_stState.bValid AND q_stState.fSocPct>=0 AND q_stState.fSocPct<=100;
_stBat.stSoh.fValue:=q_stState.fSohPct;
_stBat.stSoh.bValid:=q_stState.bValid AND q_stState.fSohPct>=0 AND q_stState.fSohPct<=100;
_stBat.fPChgMax:=SEL(q_stState.bValid,0.0,q_stState.fChargeLimitKw);
_stBat.fPDisMax:=SEL(q_stState.bValid,0.0,q_stState.fDischargeLimitKw);
_stBat.bWriteFail:=_bWriteFail;
IF NOT _fbJob.q_bBusy AND NOT _fbJob.q_bDone AND i_bEnable AND i_sIpAddr<>'' THEN
IF _bPendingWrite THEN
 _nAddress:=_nPendingAddress; _nQuantity:=_nPendingQty; _wValue:=_wPendingValue;
 _awValues[0]:=_wPendingValue; _awValues[1]:=_wPendingValue; _awValues[2]:=_wPendingValue;
 IF _nPendingQty>1 THEN _nFunction:=16; ELSE _nFunction:=6; END_IF
 _bCurrentWrite:=TRUE; _bPendingWrite:=FALSE; _bLaunch:=TRUE;
ELSIF _bReadDue THEN
 _bCurrentWrite:=FALSE;

 _nFunction:=4;
 CASE _nPoll OF
  0: _nAddress:=0; _nQuantity:=27; // 맵 v1.4: 30001~30027
  1: _nAddress:=50; _nQuantity:=40;
  2: _nAddress:=90; _nQuantity:=90;
  3:
   IF NOT i_bReadDetails THEN _nPoll:=0; _nAddress:=0; _nQuantity:=27;
   ELSE
    _nDetailChunk:=MIN(125,406-_nDetailOffset);
    _nAddress:=UINT_TO_WORD(500+500*(_nDetailRack-1)+_nDetailOffset);
    _nQuantity:=UINT_TO_WORD(_nDetailChunk);
   END_IF
 END_CASE
 _bLaunch:=TRUE;
 END_IF
END_IF
IF NOT i_bEnable THEN _nSampleSeq:=0; _nPoll:=0; _nDetailOffset:=0; _bLaunch:=FALSE; END_IF
END_METHOD

PROPERTY BatState : ST_BatState
GET
BatState:=_stBat;
END_GET
END_PROPERTY

METHOD PRIVATE M_QueueWrite : BOOL
VAR_INPUT i_nAddress : WORD; i_wValue : WORD;
 i_nQuantity : WORD; // 1 = FC06. 2~3 = FC16로 i_nAddress부터 같은 값 i_wValue를 여러 칸에 [2026-11-13]
END_VAR
q_eRequestResult := E_UpsResult.Disabled;
IF NOT GVL_PARAM.UPS_CONTROL_ENABLED OR NOT i_bWritePermit OR NOT i_bEnable THEN RETURN; END_IF
IF i_nQuantity<1 OR i_nQuantity>3 THEN q_eRequestResult := E_UpsResult.BadRequest; RETURN; END_IF
q_eRequestResult := E_UpsResult.CommUnavailable;
IF NOT q_stState.bValid THEN RETURN; END_IF
q_eRequestResult := E_UpsResult.Busy;
IF _bPendingWrite OR _bCurrentWrite AND (_fbJob.q_bBusy OR _bLaunch) THEN RETURN; END_IF
_nPendingAddress := i_nAddress; _wPendingValue := i_wValue; _nPendingQty := i_nQuantity; _bPendingWrite := TRUE;
q_eRequestResult := E_UpsResult.Accepted;
M_QueueWrite := TRUE;
END_METHOD

METHOD M_SetRackMask : BOOL
// Whole installed-rack bitmap, not an individual-rack pulse. 0 disables ALL installed racks.
VAR_INPUT i_wMask : WORD; END_VAR
IF i_nRackCount<1 OR i_nRackCount>10 THEN q_eRequestResult:=E_UpsResult.BadConfig; RETURN; END_IF
_wInstalledMask:=SHL(WORD#1,i_nRackCount)-1;
IF (i_wMask AND NOT _wInstalledMask)<>0 THEN q_eRequestResult:=E_UpsResult.BadConfig; RETURN; END_IF
M_SetRackMask:=M_QueueWrite(i_nAddress:=0,i_wValue:=i_wMask,i_nQuantity:=1);
END_METHOD

METHOD M_RequestOperation : BOOL
VAR_INPUT i_eOperation : E_EsolutionOperation; END_VAR
IF TO_INT(i_eOperation)<0 OR TO_INT(i_eOperation)>9 THEN q_eRequestResult:=E_UpsResult.Unsupported; RETURN; END_IF
M_RequestOperation:=M_QueueWrite(i_nAddress:=10,i_wValue:=SHL(WORD#1,INT_TO_UINT(TO_INT(i_eOperation))),i_nQuantity:=1);
END_METHOD

METHOD M_SetStateCmd : BOOL
VAR_INPUT i_stCmd : ST_BatCmd; END_VAR
IF _bHaveCoreCmd AND _nLastCoreCmdSeq=i_stCmd.nSeq THEN
 q_eRequestResult:=E_UpsResult.Duplicate; RETURN;
END_IF
CASE i_stCmd.eCmd OF
 // 투입·개방은 40013(랙 전체)·40014(충전)·40015(방전)를 FC16 한 번에 [1,1,1] / [0,0,0] (2026-11-12 이솔루션 답: 순서 무관, 2026-11-13 사용자 결정 2안)
 E_BatCmd.Close: M_SetStateCmd:=M_QueueWrite(i_nAddress:=INT_TO_WORD(TO_INT(E_EsolutionControl.SystemContactor)),i_wValue:=1,i_nQuantity:=3);
 E_BatCmd.Open: M_SetStateCmd:=M_QueueWrite(i_nAddress:=INT_TO_WORD(TO_INT(E_EsolutionControl.SystemContactor)),i_wValue:=0,i_nQuantity:=3);
 E_BatCmd.EStop: M_SetStateCmd:=M_SetControl(E_EsolutionControl.EmergencyShutdown,TRUE);
 E_BatCmd.Reset: M_SetStateCmd:=M_QueueWrite(i_nAddress:=30,i_wValue:=1,i_nQuantity:=1);
ELSE q_eRequestResult:=E_UpsResult.Unsupported;
END_CASE
IF M_SetStateCmd THEN _bHaveCoreCmd:=TRUE; _nLastCoreCmdSeq:=i_stCmd.nSeq; END_IF
END_METHOD

METHOD M_SetControl : BOOL
// System protocol v1.4: 0-based holding addresses, uint16 values (NOT 0x55). 하나씩 제어 (EMS command/bat 5~10)
VAR_INPUT i_eControl : E_EsolutionControl; i_bOn : BOOL; END_VAR
CASE i_eControl OF
 E_EsolutionControl.EmergencyShutdown:
  IF NOT i_bOn THEN q_eRequestResult:=E_UpsResult.Unsupported; RETURN; END_IF;
  M_SetControl:=M_QueueWrite(i_nAddress:=11,i_wValue:=1,i_nQuantity:=1);
 E_EsolutionControl.SystemContactor, E_EsolutionControl.ChargeContactor, E_EsolutionControl.DischargeContactor:
  M_SetControl:=M_QueueWrite(i_nAddress:=INT_TO_WORD(TO_INT(i_eControl)),i_wValue:=BOOL_TO_WORD(i_bOn),i_nQuantity:=1);
ELSE q_eRequestResult:=E_UpsResult.Unsupported;
END_CASE
END_METHOD

METHOD M_CheckSet : WSTRING(63)
M_CheckSet:="";
IF i_bEnable THEN
 IF i_sIpAddr='' OR i_nPort=0 THEN M_CheckSet:="TCP endpoint missing";
 ELSIF i_tReadPeriod<=T#0MS OR i_tTimeout<=T#0MS OR i_tCommTimeout<=i_tReadPeriod THEN M_CheckSet:="Invalid timing";
 END_IF
END_IF
IF i_nRackCount<1 OR i_nRackCount>10 OR i_nModuleCount<1 OR i_nModuleCount>17 THEN
 M_CheckSet:="Rack/module range";
END_IF
END_METHOD

END_FUNCTION_BLOCK

// ---- 20_Module/Ups/FB_UpsModbusJob.TcPOU
FUNCTION_BLOCK FB_UpsModbusJob
// One latched Modbus transaction. FC03/04 read, FC06 single write, FC16 block write (max 3 words, BMS 40013~40015 [2026-11-13]).
VAR_INPUT
 i_sIpAddr : STRING(15);
 i_nPort : UINT := 502;
 i_nUnitId : BYTE := 1;
 i_tTimeout : TIME := T#1S;
 i_bExecute : BOOL;
 i_bWritePermit : BOOL;
 i_nFunction : UINT;
 i_nAddress : WORD;
 i_nQuantity : WORD;
 i_wValue : WORD;
 i_awValues : ARRAY[0..2] OF WORD; // FC16 values (i_nQuantity words) [2026-11-13]
END_VAR
VAR_OUTPUT
 q_bBusy : BOOL;
 q_bDone : BOOL;
 q_bError : BOOL;
 q_nErrorId : UDINT;
 q_awData : ARRAY[0..124] OF WORD;
END_VAR
VAR
 _fbInput : FB_MBReadInputRegs;
 _fbHolding : FB_MBReadRegs;
 _fbSingle : FB_MBWriteSingleReg;
 _fbMulti : FB_MBWriteRegs; // FC16 [2026-11-13]
 _awValues : ARRAY[0..2] OF WORD;
 _bStartMulti : BOOL;
 _rtExecute : R_TRIG;
 _sIpAddr : STRING(15);
 _nPort : UINT;
 _nUnitId : BYTE;
 _tTimeout : TIME;
 _nAddress : WORD;
 _wValue : WORD;
 _nFunction : UINT;
 _nQuantity : WORD;
 _bStartInput : BOOL;
 _bStartHolding : BOOL;
 _bStartWrite : BOOL;
END_VAR

q_bDone := FALSE;
q_bError := FALSE;
_bStartInput := FALSE; _bStartHolding := FALSE; _bStartWrite := FALSE; _bStartMulti := FALSE;
_rtExecute(CLK := i_bExecute);
IF _rtExecute.Q AND NOT q_bBusy THEN
 q_nErrorId := 0;
 IF i_sIpAddr = '' OR i_nPort = 0 OR i_nQuantity = 0 OR i_nQuantity > 125 THEN
  q_bDone := TRUE; q_bError := TRUE; q_nErrorId := 16#F001;
 ELSIF (i_nFunction = 6 AND (NOT GVL_PARAM.UPS_CONTROL_ENABLED OR NOT i_bWritePermit OR i_nQuantity <> 1))
  OR (i_nFunction = 16 AND (NOT GVL_PARAM.UPS_CONTROL_ENABLED OR NOT i_bWritePermit OR i_nQuantity > 3)) THEN
  q_bDone := TRUE; q_bError := TRUE; q_nErrorId := 16#F002;
 ELSIF i_nFunction <> 3 AND i_nFunction <> 4 AND i_nFunction <> 6 AND i_nFunction <> 16 THEN
  q_bDone := TRUE; q_bError := TRUE; q_nErrorId := 16#F003;
 ELSE
  _sIpAddr:=i_sIpAddr; _nPort:=i_nPort; _nUnitId:=i_nUnitId;
  _tTimeout:=i_tTimeout; _nAddress:=i_nAddress; _wValue:=i_wValue; _awValues:=i_awValues;
  _nFunction := i_nFunction; _nQuantity := i_nQuantity; q_bBusy := TRUE;
  _bStartInput := _nFunction = 4; _bStartHolding := _nFunction = 3; _bStartWrite := _nFunction = 6;
  _bStartMulti := _nFunction = 16;
 END_IF
END_IF
// Call all instances every scan, also while disabled, to drain an in-flight transaction.
_fbInput(sIPAddr:=_sIpAddr,nTCPPort:=_nPort,nUnitID:=_nUnitId,nMBAddr:=_nAddress,nQuantity:=_nQuantity,
 cbLength:=SIZEOF(q_awData),pDestAddr:=ADR(q_awData),tTimeout:=_tTimeout,bExecute:=_bStartInput);
_fbHolding(sIPAddr:=_sIpAddr,nTCPPort:=_nPort,nUnitID:=_nUnitId,nMBAddr:=_nAddress,nQuantity:=_nQuantity,
 cbLength:=SIZEOF(q_awData),pDestAddr:=ADR(q_awData),tTimeout:=_tTimeout,bExecute:=_bStartHolding);
_fbSingle(sIPAddr:=_sIpAddr,nTCPPort:=_nPort,nUnitID:=_nUnitId,nMBAddr:=_nAddress,nValue:=_wValue,tTimeout:=_tTimeout,bExecute:=_bStartWrite);
_fbMulti(sIPAddr:=_sIpAddr,nTCPPort:=_nPort,nUnitID:=_nUnitId,nQuantity:=_nQuantity,nMBAddr:=_nAddress,
 cbLength:=WORD_TO_UDINT(_nQuantity)*2,pSrcAddr:=ADR(_awValues),tTimeout:=_tTimeout,bExecute:=_bStartMulti);
IF q_bBusy THEN
 CASE _nFunction OF
  4: IF NOT _fbInput.bBusy AND NOT _bStartInput THEN
    q_bDone := TRUE; q_bError := _fbInput.bError OR (_fbInput.cbRead <> WORD_TO_UDINT(_nQuantity)*2);
    q_nErrorId := _fbInput.nErrId; q_bBusy := FALSE; END_IF
  3: IF NOT _fbHolding.bBusy AND NOT _bStartHolding THEN
    q_bDone := TRUE; q_bError := _fbHolding.bError OR (_fbHolding.cbRead <> WORD_TO_UDINT(_nQuantity)*2);
    q_nErrorId := _fbHolding.nErrId; q_bBusy := FALSE; END_IF
  6: IF NOT _fbSingle.bBusy AND NOT _bStartWrite THEN
    q_bDone := TRUE; q_bError := _fbSingle.bError; q_nErrorId := _fbSingle.nErrId; q_bBusy := FALSE; END_IF
  16: IF NOT _fbMulti.bBusy AND NOT _bStartMulti THEN
    q_bDone := TRUE; q_bError := _fbMulti.bError; q_nErrorId := _fbMulti.nErrId; q_bBusy := FALSE; END_IF
 END_CASE
 IF q_bDone AND q_bError AND q_nErrorId = 0 THEN q_nErrorId := 16#F004; END_IF
END_IF

END_FUNCTION_BLOCK

// ---- 20_Module/Ups/F_UpsNextSeq.TcPOU
FUNCTION F_UpsNextSeq : UDINT
VAR_INPUT i_nSeq : UDINT; END_VAR

IF i_nSeq = 16#FFFFFFFF THEN F_UpsNextSeq := 1;
ELSE F_UpsNextSeq := i_nSeq + 1; END_IF

END_FUNCTION

// ---- 20_Module/Virtual/FB_MeterSim.TcPOU
FUNCTION_BLOCK FB_MeterSim EXTENDS FB_DeviceBase IMPLEMENTS I_Meter		// 가상 계측기 (시험용)
VAR_INPUT
	i_fP			: REAL;					// kW (방전 +). PRG_SimLink가 넣음
	i_fQ			: REAL;					// kvar
	i_fVPhase		: REAL := 13221.0;		// V, 상전압
	i_fHz			: REAL := 60.0;
	i_bForceInvalid	: BOOL;			// 시험: 접속점 P/Q 계측 무효 (값·통신·전압·주파수는 유지)
END_VAR
VAR
	_stMeter		: ST_MeterState;
END_VAR

PROPERTY MeterState : ST_MeterState
GET
MeterState := _stMeter;
END_GET
END_PROPERTY

METHOD M_Cycle
VAR
	k		: UINT;
END_VAR
IF M_IsReadTime() THEN		// 읽기 주기마다 응답한 것으로 봄
	M_MarkAlive();
END_IF
M_UpdateComm();

_stMeter.bComm			:= _bComm;
_stMeter.stP.fValue		:= i_fP;
_stMeter.stP.bValid		:= NOT i_bForceInvalid;
_stMeter.stQ.fValue		:= i_fQ;
_stMeter.stQ.bValid		:= NOT i_bForceInvalid;
_stMeter.stV.fValue		:= i_fVPhase;
_stMeter.stV.bValid		:= TRUE;
FOR k := 1 TO 3 DO
	_stMeter.astV[k].fValue	:= i_fVPhase;
	_stMeter.astV[k].bValid	:= TRUE;
END_FOR
_stMeter.stF.fValue		:= i_fHz;
_stMeter.stF.bValid		:= TRUE;
END_METHOD

END_FUNCTION_BLOCK

// ---- 20_Module/Driver/Sebang/FB_SebangUps.TcPOU
FUNCTION_BLOCK FB_SebangUps EXTENDS FB_DeviceBase IMPLEMENTS I_Ups

VAR_INPUT
 i_bEnable : BOOL;
 i_sIpAddr : STRING(15);
 i_nPort : UINT := 502;
 i_nUnitId : BYTE := 1;
 i_tTimeout : TIME := T#1S;
 i_bWritePermit : BOOL; // site dispatcher: config OK AND active PLC
END_VAR
VAR_OUTPUT
 q_eRequestResult : E_UpsResult;
 q_nTransportError : UDINT;
END_VAR
VAR
 _fbJob : FB_UpsModbusJob;
 _bLaunch : BOOL;
 _bCurrentWrite : BOOL;
 _bDiscardResponse : BOOL; // response started before a disable must not complete a new snapshot
 _nFunction : UINT;
 _nAddress : WORD;
 _nQuantity : WORD;
 _wValue : WORD;
 _bPendingWrite : BOOL;
 _nPendingAddress : WORD;
 _wPendingValue : WORD;
 _nPoll : UINT;
 _nCopy : UINT;
 _bReadDue : BOOL;
END_VAR

VAR_OUTPUT
 q_stRaw : ST_UpsRaw;
 q_stState : ST_UpsState;
END_VAR
VAR
 _stWork : ST_UpsRaw;
 _nSampleSeq : UDINT;
END_VAR

METHOD M_Cycle
_bReadDue := M_IsReadTime();
IF NOT i_bEnable THEN
 _bDiscardResponse:=_bDiscardResponse OR _fbJob.q_bBusy;
 _bLaunch:=FALSE;
END_IF
IF NOT i_bEnable OR NOT i_bWritePermit OR NOT GVL_PARAM.UPS_CONTROL_ENABLED THEN
 _bPendingWrite := FALSE;
 // A queued but not yet started FC06 must not survive a gate transition.
 IF _bLaunch AND _bCurrentWrite THEN _bLaunch := FALSE; END_IF
END_IF
_fbJob(i_sIpAddr:=i_sIpAddr,i_nPort:=i_nPort,i_nUnitId:=i_nUnitId,i_tTimeout:=i_tTimeout,
 i_bExecute:=_bLaunch,i_bWritePermit:=i_bWritePermit AND i_bEnable,
 i_nFunction:=_nFunction,i_nAddress:=_nAddress,i_nQuantity:=_nQuantity,i_wValue:=_wValue);
_bLaunch := FALSE;
IF _fbJob.q_bDone THEN
 q_nTransportError := _fbJob.q_nErrorId;
 IF _bCurrentWrite THEN M_MarkWriteResult(NOT _fbJob.q_bError); END_IF
END_IF

IF _fbJob.q_bDone AND _bDiscardResponse THEN
 _bDiscardResponse:=FALSE; _nPoll:=0;
ELSIF _fbJob.q_bDone AND NOT _bCurrentWrite THEN
 IF _fbJob.q_bError THEN _nPoll:=0;
 ELSE
  CASE _nPoll OF
   0: FOR _nCopy:=0 TO 34 DO _stWork.awInput[_nCopy]:=_fbJob.q_awData[_nCopy]; END_FOR
   1: FOR _nCopy:=0 TO 15 DO _stWork.awInput[_nCopy+38]:=_fbJob.q_awData[_nCopy]; END_FOR
   2: FOR _nCopy:=0 TO 11 DO _stWork.awParam[_nCopy]:=_fbJob.q_awData[_nCopy]; END_FOR
   3: FOR _nCopy:=0 TO 16 DO _stWork.awParam[_nCopy+50]:=_fbJob.q_awData[_nCopy]; END_FOR
  END_CASE
  IF _nPoll=3 THEN
   q_stRaw:=_stWork; _nSampleSeq:=F_UpsNextSeq(_nSampleSeq); M_MarkAlive(); _nPoll:=0;
  ELSE _nPoll:=_nPoll+1; END_IF
 END_IF
END_IF
M_UpdateComm();
q_stState:=F_DecodeSebangUps(q_stRaw);
q_stState.bComm:=_bComm AND i_bEnable;
q_stState.bValid:=q_stState.bComm AND _nSampleSeq<>0;
q_stState.nSampleSeq:=_nSampleSeq;
q_stState.bWriteFail:=_bWriteFail;
IF NOT _fbJob.q_bBusy AND NOT _fbJob.q_bDone AND i_bEnable AND i_sIpAddr<>'' THEN
IF _bPendingWrite THEN
 _nFunction:=6; _nAddress:=_nPendingAddress; _nQuantity:=1; _wValue:=_wPendingValue;
 _bCurrentWrite:=TRUE; _bPendingWrite:=FALSE; _bLaunch:=TRUE;
ELSIF _bReadDue THEN
 _bCurrentWrite:=FALSE;

 CASE _nPoll OF
  0: _nFunction:=4; _nAddress:=0; _nQuantity:=35;
  1: _nFunction:=4; _nAddress:=38; _nQuantity:=16;
  2: _nFunction:=3; _nAddress:=0; _nQuantity:=12;
  3: _nFunction:=3; _nAddress:=50; _nQuantity:=17;
 END_CASE
 _bLaunch:=TRUE;
 END_IF
END_IF
IF NOT i_bEnable THEN _nSampleSeq:=0; _nPoll:=0; _bLaunch:=FALSE; END_IF
END_METHOD

PROPERTY UpsState : ST_UpsState
GET
UpsState:=q_stState;
END_GET
END_PROPERTY

METHOD PRIVATE M_QueueWrite : BOOL
VAR_INPUT i_nAddress : WORD; i_wValue : WORD; END_VAR
q_eRequestResult := E_UpsResult.Disabled;
IF NOT GVL_PARAM.UPS_CONTROL_ENABLED OR NOT i_bWritePermit OR NOT i_bEnable THEN RETURN; END_IF
q_eRequestResult := E_UpsResult.CommUnavailable;
IF NOT _bComm THEN RETURN; END_IF
q_eRequestResult := E_UpsResult.Busy;
IF _bPendingWrite OR _bCurrentWrite AND (_fbJob.q_bBusy OR _bLaunch) THEN RETURN; END_IF
_nPendingAddress := i_nAddress; _wPendingValue := i_wValue; _bPendingWrite := TRUE;
q_eRequestResult := E_UpsResult.Accepted;
M_QueueWrite := TRUE;
END_METHOD

METHOD M_RequestCommand : BOOL
VAR_INPUT i_eCommand : E_UpsCommand; END_VAR
CASE i_eCommand OF
 E_UpsCommand.Reset,
 E_UpsCommand.BuzzerStop,
 E_UpsCommand.RectifierOn,
 E_UpsCommand.RectifierOff,
 E_UpsCommand.InverterOn,
 E_UpsCommand.InverterOff,
 E_UpsCommand.BbcOn,
 E_UpsCommand.BbcOff,
 E_UpsCommand.ToInverter,
 E_UpsCommand.ToBypass,
 E_UpsCommand.FloatCharge,
 E_UpsCommand.EqualCharge,
 E_UpsCommand.AutoOn,
 E_UpsCommand.AutoOff,
 E_UpsCommand.EmergencyDischarge,
 E_UpsCommand.PeriodicDischarge,
 E_UpsCommand.PulseDischarge,
 E_UpsCommand.CancelDischarge,
 E_UpsCommand.TrickleOn,
 E_UpsCommand.TrickleOff,
 E_UpsCommand.TemperatureOn,
 E_UpsCommand.TemperatureOff,
 E_UpsCommand.EcoOn,
 E_UpsCommand.EcoOff,
 E_UpsCommand.PrltOn,
 E_UpsCommand.PrltOff:
 M_RequestCommand:=M_QueueWrite(INT_TO_WORD(TO_INT(i_eCommand)),16#0055);
ELSE q_eRequestResult:=E_UpsResult.Unsupported;
END_CASE
END_METHOD

METHOD M_SetParameter : BOOL
// Explicit RAW register value only. Unresolved SOC/base-cell encodings are rejected.
VAR_INPUT i_nAddress : WORD; i_wRawValue : WORD; END_VAR
CASE i_nAddress OF
 7,8,10,50,51,52,53,54,55,56,60,61,63,64:
  M_SetParameter:=M_QueueWrite(i_nAddress,i_wRawValue);
ELSE q_eRequestResult:=E_UpsResult.Unsupported;
END_CASE
END_METHOD

METHOD M_CheckSet : WSTRING(63)
M_CheckSet:="";
IF i_bEnable THEN
 IF i_sIpAddr='' OR i_nPort=0 THEN M_CheckSet:="TCP endpoint missing";
 ELSIF i_tReadPeriod<=T#0MS OR i_tTimeout<=T#0MS OR i_tCommTimeout<=i_tReadPeriod THEN M_CheckSet:="Invalid timing";
 END_IF
END_IF
END_METHOD

END_FUNCTION_BLOCK

// ---- 20_Module/Driver/Sebang/F_DecodeSebangUps.TcPOU
FUNCTION F_DecodeSebangUps : ST_UpsState
VAR_INPUT i_stRaw : ST_UpsRaw; END_VAR
VAR n : UINT; END_VAR

// UPS Metering Data 주소 순서
F_DecodeSebangUps.fInputVoltageRV := WORD_TO_REAL(i_stRaw.awInput[0])*0.1; // 0. 입력 선간 전압 R (V)
F_DecodeSebangUps.fInputVoltageSV := WORD_TO_REAL(i_stRaw.awInput[1])*0.1; // 1. 입력 선간 전압 S (V)
F_DecodeSebangUps.fInputVoltageTV := WORD_TO_REAL(i_stRaw.awInput[2])*0.1; // 2. 입력 선간 전압 T (V)
F_DecodeSebangUps.fInputFrequencyHz := WORD_TO_REAL(i_stRaw.awInput[3])*0.1; // 3. 입력 주파수 (Hz)
F_DecodeSebangUps.fInputCurrentRA := WORD_TO_REAL(i_stRaw.awInput[4])*0.1; // 4. 입력 전류 R (A)
F_DecodeSebangUps.fInputCurrentSA := WORD_TO_REAL(i_stRaw.awInput[5])*0.1; // 5. 입력 전류 S (A)
F_DecodeSebangUps.fInputCurrentTA := WORD_TO_REAL(i_stRaw.awInput[6])*0.1; // 6. 입력 전류 T (A)
F_DecodeSebangUps.fInverterVoltageRV := WORD_TO_REAL(i_stRaw.awInput[7])*0.1; // 7. 인버터 선간 전압 R (V)
F_DecodeSebangUps.fInverterVoltageSV := WORD_TO_REAL(i_stRaw.awInput[8])*0.1; // 8. 인버터 선간 전압 S (V)
F_DecodeSebangUps.fInverterVoltageTV := WORD_TO_REAL(i_stRaw.awInput[9])*0.1; // 9. 인버터 선간 전압 T (V)
F_DecodeSebangUps.fInverterCurrentRA := WORD_TO_REAL(i_stRaw.awInput[10])*0.1; // 10. 인버터 전류 R (A)
F_DecodeSebangUps.fInverterCurrentSA := WORD_TO_REAL(i_stRaw.awInput[11])*0.1; // 11. 인버터 전류 S (A)
F_DecodeSebangUps.fInverterCurrentTA := WORD_TO_REAL(i_stRaw.awInput[12])*0.1; // 12. 인버터 전류 T (A)
F_DecodeSebangUps.fBypassVoltageRV := WORD_TO_REAL(i_stRaw.awInput[13])*0.1; // 13. 바이패스 선간 전압 R (V)
F_DecodeSebangUps.fBypassVoltageSV := WORD_TO_REAL(i_stRaw.awInput[14])*0.1; // 14. 바이패스 선간 전압 S (V)
F_DecodeSebangUps.fBypassVoltageTV := WORD_TO_REAL(i_stRaw.awInput[15])*0.1; // 15. 바이패스 선간 전압 T (V)
F_DecodeSebangUps.fBypassFrequencyHz := WORD_TO_REAL(i_stRaw.awInput[16])*0.1; // 16. 바이패스 주파수 (Hz)
F_DecodeSebangUps.fOutputVoltageRV := WORD_TO_REAL(i_stRaw.awInput[17])*0.1; // 17. 출력 선간 전압 R (V)
F_DecodeSebangUps.fOutputVoltageSV := WORD_TO_REAL(i_stRaw.awInput[18])*0.1; // 18. 출력 선간 전압 S (V)
F_DecodeSebangUps.fOutputVoltageTV := WORD_TO_REAL(i_stRaw.awInput[19])*0.1; // 19. 출력 선간 전압 T (V)
F_DecodeSebangUps.fOutputFrequencyHz := WORD_TO_REAL(i_stRaw.awInput[20])*0.1; // 20. 출력 주파수 (Hz)
F_DecodeSebangUps.fOutputCurrentRA := WORD_TO_REAL(i_stRaw.awInput[21])*0.1; // 21. 출력 전류 R (A)
F_DecodeSebangUps.fOutputCurrentSA := WORD_TO_REAL(i_stRaw.awInput[22])*0.1; // 22. 출력 전류 S (A)
F_DecodeSebangUps.fOutputCurrentTA := WORD_TO_REAL(i_stRaw.awInput[23])*0.1; // 23. 출력 전류 T (A)
F_DecodeSebangUps.fDcLinkVoltageV := F_UpsSignedWord(i_stRaw.awInput[24])*0.1; // 24. DC 링크 전압 (V)
F_DecodeSebangUps.fDcLinkHighVoltageV := F_UpsSignedWord(i_stRaw.awInput[25])*0.1; // 25. DC 링크 상단 전압 (V)
F_DecodeSebangUps.fDcLinkLowVoltageV := F_UpsSignedWord(i_stRaw.awInput[26])*0.1; // 26. DC 링크 하단 전압 (V)
F_DecodeSebangUps.fBatteryVoltageV := F_UpsSignedWord(i_stRaw.awInput[27])*0.1; // 27. 배터리 전압 (V)
F_DecodeSebangUps.fBatteryCurrentA := F_UpsSignedWord(i_stRaw.awInput[28])*0.1; // 28. 배터리 전류 (A)
F_DecodeSebangUps.fMpiCurrentAA := F_UpsSignedWord(i_stRaw.awInput[29])*0.1; // 29. MPI A상 전류 (A)
F_DecodeSebangUps.fMpiCurrentBA := F_UpsSignedWord(i_stRaw.awInput[30])*0.1; // 30. MPI B상 전류 (A)
F_DecodeSebangUps.fMpiCurrentCA := F_UpsSignedWord(i_stRaw.awInput[31])*0.1; // 31. MPI C상 전류 (A)
F_DecodeSebangUps.fInputApparentPowerKva := F_UpsSignedWord(i_stRaw.awInput[32])*0.1; // 32. 입력 피상 전력 (kVA)
F_DecodeSebangUps.fOutputApparentPowerKva := F_UpsSignedWord(i_stRaw.awInput[33])*0.1; // 33. 출력 피상 전력 (kVA)
F_DecodeSebangUps.fOutputActivePowerKw := F_UpsSignedWord(i_stRaw.awInput[34])*0.1; // 34. 출력 유효 전력 (kW)
F_DecodeSebangUps.fTemperature1C := F_UpsSignedWord(i_stRaw.awInput[38])*0.1; // 38. 온도 1 (℃)
F_DecodeSebangUps.fTemperature2C := F_UpsSignedWord(i_stRaw.awInput[39])*0.1; // 39. 온도 2 (℃)
F_DecodeSebangUps.fTemperature3C := F_UpsSignedWord(i_stRaw.awInput[40])*0.1; // 40. 온도 3 (℃)
F_DecodeSebangUps.fTemperature4C := F_UpsSignedWord(i_stRaw.awInput[41])*0.1; // 41. 온도 4 (℃)
F_DecodeSebangUps.fTemperature5C := F_UpsSignedWord(i_stRaw.awInput[42])*0.1; // 42. 온도 5 (℃)
F_DecodeSebangUps.fBatteryRoomTemperatureC := F_UpsSignedWord(i_stRaw.awInput[43])*0.1; // 43. 온도 6 / 배터리실 온도 (℃)
F_DecodeSebangUps.wInputAlarm := i_stRaw.awInput[44]; // 44. 입력 알람
F_DecodeSebangUps.wRectAlarm := i_stRaw.awInput[45]; // 45. 정류기 알람
F_DecodeSebangUps.wBbcAlarm := i_stRaw.awInput[46]; // 46. 배터리 컨버터 알람
F_DecodeSebangUps.wOutputAlarm := i_stRaw.awInput[47]; // 47. 출력 알람
F_DecodeSebangUps.wInverterAlarm := i_stRaw.awInput[48]; // 48. 인버터 알람
F_DecodeSebangUps.wBypassAlarm := i_stRaw.awInput[49]; // 49. 바이패스 알람
F_DecodeSebangUps.wStatus1 := i_stRaw.awInput[50]; // 50. 상태 워드 1
F_DecodeSebangUps.wStatus2 := i_stRaw.awInput[51]; // 51. 상태 워드 2
F_DecodeSebangUps.fHmiVersion := WORD_TO_REAL(i_stRaw.awInput[52])*0.1; // 52. HMI 버전
F_DecodeSebangUps.fDspVersion := WORD_TO_REAL(i_stRaw.awInput[53])*0.1; // 53. DSP 버전

F_DecodeSebangUps.nBatMode := WORD_TO_UINT(SHR(i_stRaw.awInput[50],8) AND 16#0007);
F_DecodeSebangUps.bRectOn := i_stRaw.awInput[45].11;
F_DecodeSebangUps.bRectNormal := i_stRaw.awInput[45].12;
F_DecodeSebangUps.bBbcOn := i_stRaw.awInput[46].12;
F_DecodeSebangUps.bBbcNormal := i_stRaw.awInput[46].13;
F_DecodeSebangUps.bInverterOn := i_stRaw.awInput[48].6;
F_DecodeSebangUps.bInverterNormal := i_stRaw.awInput[48].14;
F_DecodeSebangUps.bOnBypass := i_stRaw.awInput[48].12;
F_DecodeSebangUps.bOnInverter := i_stRaw.awInput[48].13;
F_DecodeSebangUps.bTemperatureEnabled := i_stRaw.awInput[51].2;
F_DecodeSebangUps.bBmsMinor := i_stRaw.awInput[51].10;
F_DecodeSebangUps.bBmsMajor := i_stRaw.awInput[51].11;
F_DecodeSebangUps.bEmergencyStop := i_stRaw.awInput[50].0;
FOR n:=0 TO 7 DO F_DecodeSebangUps.awAlarmStatus[n]:=i_stRaw.awInput[n+44]; END_FOR

END_FUNCTION

// ---- 20_Module/Common/FB_RuleBit.TcPOU
FUNCTION_BLOCK FB_RuleBit EXTENDS FB_ModuleBase IMPLEMENTS I_ProtectionRule, I_OutputRule		// 디지털 접점 하나 → 조건 (화재·연기·비상정지·문 열림 등). 보호 규칙·출력 규칙 어느 쪽으로도 등록
VAR_INPUT
	i_ipAux			: I_AuxDevice;		// 읽을 보조 장비 (선언 때 지정)
	i_nPoint		: UINT;				// 디지털 입력 점 번호
	i_stSet			: ST_RuleBitSet;	// 설정: b접점, 통신 끊김 시 조건 (MAIN이 GVL_PERSIST.g_stModuleSet 칸을 매 스캔 넘김. 안 넘기면 기본값)
END_VAR
VAR
	_bCond			: BOOL;
END_VAR

METHOD M_Evaluate : BOOL		// 보호 규칙으로 판단 (범위·대상과 관계없이 접점 하나)
VAR_INPUT
	i_stView	: ST_ProtView;
END_VAR
M_Evaluate := M_Check(i_fThreshold := i_stView.fThreshold);
END_METHOD

METHOD M_Check : BOOL		// 출력 규칙으로 판단. 보호 판단도 이것을 씀
VAR_INPUT
	i_fThreshold	: REAL;			// 안 씀
END_VAR
IF i_ipAux = 0 THEN
	_bCond := FALSE;
ELSIF NOT i_ipAux.Comm THEN
	_bCond := i_stSet.bOnCommLoss;
ELSE
	_bCond := i_ipAux.M_GetBit(i_nPoint) XOR i_stSet.bInvert;
END_IF
M_Check := _bCond;
END_METHOD

END_FUNCTION_BLOCK

// ---- 20_Module/Driver/Autonics/FB_AutonicsThd.TcPOU
FUNCTION_BLOCK FB_AutonicsThd EXTENDS FB_DeviceBase IMPLEMENTS I_AuxDevice		// 오토닉스 THD 온습도계 (Modbus RTU, 한 줄에 국번 1..n), 읽기 전용
(* ---------------------------------------------------------------
   기반: Helios FB_ThdAutonics_Chain (PRG_Sensor에서 쓰던 것). 동작만 옮기고 PmsStd 드라이버 형식으로 다시 씀. 2026-11-09
   통신: 시리얼 단자(EL6022 채널 하나, 사용자 2026-11-09 회사 표준)를 ModbusRtuMaster_KL6x22B로. 단자 연결(InData·OutData)은 XAE I/O 화면에서 사람이 함
   읽기: 읽기 주기마다 센서 하나씩 돌아가며 Input Register(FC4)
     @MAP IR 0 S16 0.01 ℃  온도
     @MAP IR 1 S16 0.01 %  습도
   점 (I_AuxDevice)
     AI 2n-1 = 센서 n 온도 (℃), AI 2n = 센서 n 습도 (%). 센서 n이 i_tCommTimeout 동안 응답 없으면 bValid FALSE
     DI n    = 센서 n 통신 이상 (TRUE = 이상. Helios SensorStatus 1과 같음)
   센서는 GVL_PARAM.AUX_AI_MAX / 2개까지. 쓰기(DO·AO) 없음
   맵 미확보: Helios 현장 기종 기준. 실제 기종이 정해지면 주소·배율 확인
   --------------------------------------------------------------- *)
VAR_INPUT
	i_bEnable		: BOOL;					// FALSE면 통신하지 않음 (장비 미설치)
	i_nSensorCount	: UINT := 1;			// 국번 1..n 연속 (1..SENSOR_MAX)
	i_tTimeout		: TIME := T#1S;			// 응답 기다림 (Helios 5 s)
END_VAR
VAR
	_fbRtu			: ModbusRtuMaster_KL6x22B;
	_awRaw			: ARRAY[0..1] OF WORD;
	_bReadDue		: BOOL;					// 읽을 때가 됨 (매 스캔 M_IsReadTime)
	_bReading		: BOOL;
	_nUnit			: UINT;					// 지금 읽는 국번
	_nCount			: UINT;					// 쓰는 센서 수 (범위로 자른 i_nSensorCount)
	_afTemp			: ARRAY[1..SENSOR_MAX] OF REAL;
	_afHum			: ARRAY[1..SENSOR_MAX] OF REAL;
	_abReadOk		: ARRAY[1..SENSOR_MAX] OF BOOL;	// 이번 스캔에 응답 받음
	_abEverOk		: ARRAY[1..SENSOR_MAX] OF BOOL;	// 한 번이라도 응답 받음
	_abSensorOk		: ARRAY[1..SENSOR_MAX] OF BOOL;	// 센서 통신 정상
	_atonLoss		: ARRAY[1..SENSOR_MAX] OF TON;
	_nIdx			: UINT;
END_VAR
VAR CONSTANT
	SENSOR_MAX		: UINT := GVL_PARAM.AUX_AI_MAX / 2;
END_VAR

METHOD M_Cycle
_nCount := LIMIT(1, i_nSensorCount, SENSOR_MAX);

_bReadDue := M_IsReadTime();
IF NOT _bReading THEN
	IF i_bEnable AND _bReadDue THEN
		IF _nUnit >= _nCount THEN _nUnit := 1; ELSE _nUnit := _nUnit + 1; END_IF
		_fbRtu.ReadInputRegs(UnitID := UINT_TO_BYTE(_nUnit), Quantity := 2, MBAddr := 0,
			cbLength := SIZEOF(_awRaw), pMemoryAddr := ADR(_awRaw), Timeout := i_tTimeout, Execute := TRUE);
		_bReading := TRUE;
	END_IF
ELSE
	_fbRtu.ReadInputRegs(Execute := FALSE);	// 시작한 읽기는 끝까지 부름 (Helios와 같음)
	IF NOT _fbRtu.BUSY THEN
		IF NOT _fbRtu.Error AND i_bEnable THEN
			_afTemp[_nUnit]		:= INT_TO_REAL(WORD_TO_INT(_awRaw[0])) * 0.01;	// @MAP IR 0 S16 0.01 ℃
			_afHum[_nUnit]		:= INT_TO_REAL(WORD_TO_INT(_awRaw[1])) * 0.01;	// @MAP IR 1 S16 0.01 %
			_abReadOk[_nUnit]	:= TRUE;
			_abEverOk[_nUnit]	:= TRUE;
			M_MarkAlive();
		END_IF
		_bReading := FALSE;
	END_IF
END_IF

FOR _nIdx := 1 TO SENSOR_MAX DO
	_atonLoss[_nIdx](IN := NOT _abReadOk[_nIdx], PT := i_tCommTimeout);
	_abSensorOk[_nIdx]	:= i_bEnable AND _nIdx <= _nCount AND _abEverOk[_nIdx] AND NOT _atonLoss[_nIdx].Q;
	_abReadOk[_nIdx]	:= FALSE;
END_FOR
M_UpdateComm();
END_METHOD

METHOD M_GetBit : BOOL		// DI n = 센서 n 통신 이상
VAR_INPUT
	i_nPoint	: UINT;
END_VAR
IF i_nPoint >= 1 AND i_nPoint <= _nCount THEN
	M_GetBit := NOT _abSensorOk[i_nPoint];
END_IF
END_METHOD

METHOD M_GetValue : ST_Val		// AI 2n-1 = 센서 n 온도 (℃), AI 2n = 센서 n 습도 (%)
VAR_INPUT
	i_nPoint	: UINT;
END_VAR
VAR
	nSensor		: UINT;
END_VAR
nSensor := (i_nPoint + 1) / 2;
IF i_nPoint >= 1 AND nSensor <= _nCount THEN
	M_GetValue.fValue := SEL(i_nPoint MOD 2 = 1, _afHum[nSensor], _afTemp[nSensor]);
	M_GetValue.bValid := _abSensorOk[nSensor];
END_IF
END_METHOD

METHOD M_SetBit		// 출력 없음
VAR_INPUT
	i_nPoint	: UINT;
	i_bValue	: BOOL;
END_VAR
;
END_METHOD

METHOD M_SetValue		// 출력 없음
VAR_INPUT
	i_nPoint	: UINT;
	i_fValue	: REAL;
END_VAR
;
END_METHOD

PROPERTY Comm : BOOL
GET
Comm := _bComm AND i_bEnable;
END_GET
END_PROPERTY

END_FUNCTION_BLOCK

// ---- 20_Module/Driver/LS/FB_LsImd1000.TcPOU
FUNCTION_BLOCK FB_LsImd1000 EXTENDS FB_DeviceBase IMPLEMENTS I_AuxDevice		// LS IMD1000 절연감시장치(IMD) (Modbus TCP, RS485 게이트웨이 경유), 읽기 전용
(* ---------------------------------------------------------------
   기반: MESSIS(TC2) FB_LsIMD1000. 주소는 LS 맵으로 고침. 2026-11-09
   맵: 인터페이스\(MM-20210721) IMD1000 Modbus-Setting_v1_0_0.pdf (장비는 RS485 RTU 전용 → 현장은 RS485-TCP 게이트웨이, 사용자 결정)
   읽기 (프로토콜 주소, 0 기준 = 맵 Addr 열)
     측정: Input Register(FC4) 199부터 36개 (MESSIS와 같은 범위)
       @MAP IR 206 U16  기기 DI 입력 상태
       @MAP IR 209 U16  자가진단 Error #2
       @MAP IR 210 U16  절연저항 alarm 상태
       @MAP IR 211 U16  기기 & 계통 연결 상태
       @MAP IR 215 U16  Self Test 진행 상태
       @MAP IR 224~225 F32(앞 = 상위)  절연저항 kΩ
       MESSIS는 223~224를 읽어 한 칸 어긋나 있었다(223 = 커패시턴스 상태). 상위 워드가 맞아 값은 거의 같게 보였음
     설정: Holding Register(FC3) 40부터 8개, 측정 SET_EVERY번에 한 번
       @MAP HR 40~41 U32(앞 = 상위)  Ins. Alarm Pick-up kΩ
       @MAP HR 46~47 U32  Pre Alarm#1 Pick-up kΩ
   점 (I_AuxDevice). DI 2는 Bender ISO685 드라이버와 같은 "보호용 경보"
     AI 1 절연저항, 2 Ins. Alarm 설정값, 3 Pre Alarm#1 설정값
     DI 1 경고 (Pre#1 OR Pre#2), 2 절연 경보 (Ins. Alarm), 3 시험 중, 4 사전경고 (Pre#3), 5 기기 고장 (자가진단·Device), 6 계통 연결 이상, 7 접지(PE) 연결 이상
   쓰기 없음 (릴레이·Self Test 제어는 하지 않음)
   --------------------------------------------------------------- *)
VAR_INPUT
	i_bEnable		: BOOL;					// FALSE면 통신하지 않음 (장비 미설치)
	i_sIpAddr		: STRING(15);			// 게이트웨이 주소
	i_nPort			: UINT := 502;
	i_nUnitId		: BYTE := 1;			// IMD1000 국번 (장비 초기값 1)
	i_tTimeout		: TIME := T#1S;
END_VAR
VAR_OUTPUT
	q_stState		: ST_LsImd1000State;	// 읽은 값 (보고 매핑 FB_RptLsImd1000이 씀)
END_VAR
VAR
	_fbIr			: FB_MBReadInputRegs;	// 측정 (FC4)
	_fbHr			: FB_MBReadRegs;		// 설정 (FC3)
	_awIr			: ARRAY[0..35] OF WORD;	// IR 199..234
	_awSet			: ARRAY[0..7] OF WORD;	// HR 40..47
	_bReadDue		: BOOL;					// 읽을 때가 됨 (매 스캔 M_IsReadTime)
	_bReading		: BOOL;
	_bSetBlock		: BOOL;					// 이번 읽기가 설정 영역
	_bBusy			: BOOL;
	_bError			: BOOL;
	_nReadCnt		: UINT;					// 0이면 설정 영역을 읽음 (부팅 직후 먼저)
	_bMeasOk		: BOOL;					// 측정 영역을 한 번 이상 읽음
END_VAR
VAR CONSTANT
	IR_ADDR			: UINT := 199;
	IR_QTY			: UINT := 36;
	SET_ADDR		: UINT := 40;
	SET_QTY			: UINT := 8;
	SET_EVERY		: UINT := 10;			// 설정 영역은 읽기 10번에 한 번
END_VAR

ACTION A_MapMeas:
q_stState.wDiState		:= _awIr[7];		// @MAP IR 206
q_stState.wSelfDiag		:= _awIr[10];		// @MAP IR 209
q_stState.wAlarm		:= _awIr[11];		// @MAP IR 210
q_stState.wConnect		:= _awIr[12];		// @MAP IR 211
q_stState.wSelfTest		:= _awIr[16];		// @MAP IR 215
q_stState.fInsulation	:= F_WordsToReal(i_wHigh := _awIr[25], i_wLow := _awIr[26]);	// @MAP IR 224(상위)·225(하위) F32 kΩ
_bMeasOk := TRUE;
END_ACTION

ACTION A_MapSet:
q_stState.nInsPickup	:= SHL(WORD_TO_UDINT(_awSet[0]), 16) OR WORD_TO_UDINT(_awSet[1]);	// @MAP HR 40~41 U32
q_stState.nPre1Pickup	:= SHL(WORD_TO_UDINT(_awSet[6]), 16) OR WORD_TO_UDINT(_awSet[7]);	// @MAP HR 46~47 U32
q_stState.bSetValid		:= TRUE;
END_ACTION

METHOD M_Cycle
_bReadDue := M_IsReadTime();
IF NOT _bReading THEN
	IF i_bEnable AND i_sIpAddr <> '' AND _bReadDue THEN
		_bSetBlock := _nReadCnt = 0;
		IF _bSetBlock THEN
			_fbHr(sIPAddr := i_sIpAddr, nTCPPort := i_nPort, nUnitID := i_nUnitId,
				nQuantity := SET_QTY, nMBAddr := SET_ADDR, cbLength := SIZEOF(_awSet),
				pDestAddr := ADR(_awSet), tTimeout := i_tTimeout, bExecute := TRUE);
		ELSE
			_fbIr(sIPAddr := i_sIpAddr, nTCPPort := i_nPort, nUnitID := i_nUnitId,
				nQuantity := IR_QTY, nMBAddr := IR_ADDR, cbLength := SIZEOF(_awIr),
				pDestAddr := ADR(_awIr), tTimeout := i_tTimeout, bExecute := TRUE);
		END_IF
		_bReading := TRUE;
	END_IF
ELSE
	IF _bSetBlock THEN
		_fbHr(bExecute := FALSE);
		_bBusy := _fbHr.bBusy;
		_bError := _fbHr.bError;
	ELSE
		_fbIr(bExecute := FALSE);
		_bBusy := _fbIr.bBusy;
		_bError := _fbIr.bError;
	END_IF
	IF NOT _bBusy THEN
		IF NOT _bError AND i_bEnable THEN
			IF _bSetBlock THEN
				A_MapSet();
			ELSE
				A_MapMeas();
			END_IF
			M_MarkAlive();
		END_IF
		_nReadCnt := (_nReadCnt + 1) MOD SET_EVERY;
		_bReading := FALSE;
	END_IF
END_IF
M_UpdateComm();
q_stState.bValid := Comm AND _bMeasOk;
END_METHOD

METHOD M_GetBit : BOOL		// DI 1..7 (머리 주석). 통신 이상이면 FALSE (규칙 FB_RuleBit은 Comm으로 따로 판단)
VAR_INPUT
	i_nPoint	: UINT;
END_VAR
IF q_stState.bValid THEN
	CASE i_nPoint OF
		1: M_GetBit := q_stState.wAlarm.1 OR q_stState.wAlarm.2;
		2: M_GetBit := q_stState.wAlarm.0;
		3: M_GetBit := q_stState.wSelfTest = 1 OR q_stState.wDiState.0 OR q_stState.wDiState.1;
		4: M_GetBit := q_stState.wAlarm.3;
		5: M_GetBit := (q_stState.wSelfDiag AND 16#0007) <> 0 OR q_stState.wConnect.1;
		6: M_GetBit := q_stState.wConnect.2;
		7: M_GetBit := q_stState.wConnect.0;
	END_CASE
END_IF
END_METHOD

METHOD M_GetValue : ST_Val		// AI 1 절연저항 kΩ, 2 Ins. Alarm 설정값 kΩ, 3 Pre Alarm#1 설정값 kΩ
VAR_INPUT
	i_nPoint	: UINT;
END_VAR
CASE i_nPoint OF
	1:
		M_GetValue.fValue := q_stState.fInsulation;
		M_GetValue.bValid := q_stState.bValid;
	2:
		M_GetValue.fValue := UDINT_TO_REAL(q_stState.nInsPickup);
		M_GetValue.bValid := q_stState.bValid AND q_stState.bSetValid;
	3:
		M_GetValue.fValue := UDINT_TO_REAL(q_stState.nPre1Pickup);
		M_GetValue.bValid := q_stState.bValid AND q_stState.bSetValid;
END_CASE
END_METHOD

METHOD M_SetBit		// 출력 없음
VAR_INPUT
	i_nPoint	: UINT;
	i_bValue	: BOOL;
END_VAR
;
END_METHOD

METHOD M_SetValue		// 출력 없음
VAR_INPUT
	i_nPoint	: UINT;
	i_fValue	: REAL;
END_VAR
;
END_METHOD

PROPERTY Comm : BOOL
GET
Comm := _bComm AND i_bEnable;
END_GET
END_PROPERTY

END_FUNCTION_BLOCK

// ---- 20_Module/Common/F_WordsToReal.TcPOU
FUNCTION F_WordsToReal : REAL		// 레지스터 2개(IEEE754 float)를 REAL로. 앞 레지스터 = 상위 워드. 숫자가 아니면(NaN·무한) 0
(* 기반: Helios FNC_OLD_IEEE754·FNC_TO_IEEE754 (Bender ISO685, ACURA3700에서 앞 레지스터가 상위 워드). 2026-11-09 *)
VAR_INPUT
	i_wHigh		: WORD;		// 앞 레지스터 (상위 16비트)
	i_wLow		: WORD;		// 뒤 레지스터 (하위 16비트)
END_VAR
VAR
	dwRaw		: DWORD;
	fValue		: REAL;
END_VAR

dwRaw := SHL(WORD_TO_DWORD(i_wHigh), 16) OR WORD_TO_DWORD(i_wLow);
IF (dwRaw AND 16#7F800000) = 16#7F800000 THEN	// 지수부가 모두 1 = NaN·무한
	F_WordsToReal := 0.0;
ELSE
	MEMCPY(destAddr := ADR(fValue), srcAddr := ADR(dwRaw), n := 4);
	F_WordsToReal := fValue;
END_IF

END_FUNCTION

// ---- 20_Module/Driver/Rootech/FB_RootechAcuraIo.TcPOU
FUNCTION_BLOCK FB_RootechAcuraIo EXTENDS FB_DeviceBase IMPLEMENTS I_AuxDevice		// 루텍 ACURA3700 원격 I/O (Modbus TCP): 접점 입력·아날로그 입력 읽기 전용
(* ---------------------------------------------------------------
   기반: Helios FB_ACURA3700. Helios는 이 장치의 DI로 화재(열)·연기·가스 감지기 접점을 받았다. 동작만 옮기고 PmsStd 형식으로 다시 씀. 2026-11-09
   모듈 배치 (Helios와 같음, 물리 순서대로 모듈마다 레지스터 100개):
     DIO 모듈 = i_nStartAddr,  AI 모듈 = i_nStartAddr + 100.  Holding Register(FC3)
   읽기: 읽기 주기마다 DIO와 AI를 번갈아
     @MAP HR start+4..11   U16 -  DI ch1..8 상태 (0 = 꺼짐)
     @MAP HR start+16..17  U16 -  DO ch1..2 상태
     @MAP HR start+122..133 F32(앞 = 상위) -  AI ch1..6 변환값
   점 (I_AuxDevice)
     DI 1..8 = 접점 입력 ch1..8,  DI 9..10 = DO ch1..2 상태
     AI 1..6 = 아날로그 입력 ch1..6 변환값 (장치에 설정한 단위)
   쓰기(DO·AO) 없음
   맵 미확보: Helios 현장 기준. 실제 모듈 구성·주소는 현장에서 확인
   --------------------------------------------------------------- *)
VAR_INPUT
	i_bEnable		: BOOL;					// FALSE면 통신하지 않음 (장비 미설치)
	i_sIpAddr		: STRING(15);
	i_nPort			: UINT := 502;
	i_nUnitId		: BYTE := 1;
	i_nStartAddr	: UINT := 12100;		// 첫 모듈(DIO) 시작 주소
	i_tTimeout		: TIME := T#1S;
END_VAR
VAR
	_fbMbRead		: FB_MBReadRegs;
	_awDio			: ARRAY[0..41] OF WORD;
	_awAi			: ARRAY[0..45] OF WORD;
	_bReadDue		: BOOL;					// 읽을 때가 됨 (매 스캔 M_IsReadTime)
	_bReading		: BOOL;
	_bReadAi		: BOOL;					// 이번 읽기가 AI 모듈
	_abDi			: ARRAY[1..10] OF BOOL;
	_afAi			: ARRAY[1..6] OF REAL;
	_bDioOk			: BOOL;					// DIO 모듈을 한 번이라도 읽음
	_bAiOk			: BOOL;					// AI 모듈을 한 번이라도 읽음
	_nIdx			: UINT;
END_VAR

ACTION A_MapDio:
FOR _nIdx := 1 TO 8 DO
	_abDi[_nIdx] := _awDio[_nIdx + 3] <> 0;		// @MAP HR start+4..11 U16 DI ch1..8
END_FOR
_abDi[9]	:= _awDio[16] <> 0;					// @MAP HR start+16 U16 DO ch1 상태
_abDi[10]	:= _awDio[17] <> 0;					// @MAP HR start+17 U16 DO ch2 상태
END_ACTION

ACTION A_MapAi:
FOR _nIdx := 1 TO 6 DO
	_afAi[_nIdx] := F_WordsToReal(i_wHigh := _awAi[20 + 2 * _nIdx], i_wLow := _awAi[21 + 2 * _nIdx]);	// @MAP HR start+122+2(n-1) F32 AI chn
END_FOR
END_ACTION

METHOD M_Cycle
_bReadDue := M_IsReadTime();
IF NOT _bReading THEN
	IF i_bEnable AND i_sIpAddr <> '' AND _bReadDue THEN
		_bReadAi := NOT _bReadAi;
		IF _bReadAi THEN
			_fbMbRead(sIPAddr := i_sIpAddr, nTCPPort := i_nPort, nUnitID := i_nUnitId,
				nQuantity := 46, nMBAddr := i_nStartAddr + 100, cbLength := SIZEOF(_awAi),
				pDestAddr := ADR(_awAi), tTimeout := i_tTimeout, bExecute := TRUE);
		ELSE
			_fbMbRead(sIPAddr := i_sIpAddr, nTCPPort := i_nPort, nUnitID := i_nUnitId,
				nQuantity := 42, nMBAddr := i_nStartAddr, cbLength := SIZEOF(_awDio),
				pDestAddr := ADR(_awDio), tTimeout := i_tTimeout, bExecute := TRUE);
		END_IF
		_bReading := TRUE;
	END_IF
ELSE
	_fbMbRead(bExecute := FALSE);
	IF NOT _fbMbRead.bBusy THEN
		IF NOT _fbMbRead.bError AND i_bEnable THEN
			IF _bReadAi THEN
				A_MapAi();
				_bAiOk := TRUE;
			ELSE
				A_MapDio();
				_bDioOk := TRUE;
			END_IF
			M_MarkAlive();
		END_IF
		_bReading := FALSE;
	END_IF
END_IF
M_UpdateComm();
END_METHOD

METHOD M_GetBit : BOOL		// DI 1..8 = 접점 입력, 9..10 = DO 상태. 통신 이상이면 FALSE (규칙 FB_RuleBit은 Comm으로 따로 판단)
VAR_INPUT
	i_nPoint	: UINT;
END_VAR
IF i_nPoint >= 1 AND i_nPoint <= 10 AND Comm AND _bDioOk THEN
	M_GetBit := _abDi[i_nPoint];
END_IF
END_METHOD

METHOD M_GetValue : ST_Val		// AI 1..6 = 아날로그 입력 변환값
VAR_INPUT
	i_nPoint	: UINT;
END_VAR
IF i_nPoint >= 1 AND i_nPoint <= 6 THEN
	M_GetValue.fValue := _afAi[i_nPoint];
	M_GetValue.bValid := Comm AND _bAiOk;
END_IF
END_METHOD

METHOD M_SetBit		// 출력 없음 (DO는 읽기만)
VAR_INPUT
	i_nPoint	: UINT;
	i_bValue	: BOOL;
END_VAR
;
END_METHOD

METHOD M_SetValue		// 출력 없음
VAR_INPUT
	i_nPoint	: UINT;
	i_fValue	: REAL;
END_VAR
;
END_METHOD

PROPERTY Comm : BOOL
GET
Comm := _bComm AND i_bEnable;
END_GET
END_PROPERTY

END_FUNCTION_BLOCK

// ---- 20_Module/Driver/ITGuard/FB_ItGuardIeSx.TcPOU
FUNCTION_BLOCK FB_ItGuardIeSx EXTENDS FB_DeviceBase IMPLEMENTS I_AuxDevice		// ITGuard(이노튜브) IE-SX 이더넷 온습도계 (Modbus TCP), 읽기 전용
(* ---------------------------------------------------------------
   기반: MESSIS TC3 FB_IE_SX (광주첨단공장). 동작만 옮기고 PmsStd 형식으로 다시 씀. 2026-11-09
   읽기: Input Register(FC4) 0부터 5개 (MESSIS와 같음, Unit ID 1)
     @MAP IR 0  U16  mode
     @MAP IR 1  S16  센서1 = 온도 × 0.01 ℃
     @MAP IR 2  S16  센서2 = 습도 × 0.01 %
     @MAP IR 3·4 S16  센서3·4 (프로브 없으면 32767)
   2026-11-09 PC에서 읽어 확인: [0, 2418, 3545, 32767, 32767] → 24.18 ℃, 35.45 %
   센서 값 32767 = 프로브 없음으로 보고 무효 처리 (센서3·4가 비었을 때 이 값)
   점 (I_AuxDevice): AI 1 온도, AI 2 습도, DI 1 값 이상(통신 정상인데 프로브 무효)
   통신 이상: 응답 없이 i_tCommTimeout(기본 10초, MESSIS는 30초)
   쓰기 없음
   --------------------------------------------------------------- *)
VAR_INPUT
	i_bEnable		: BOOL;					// FALSE면 통신하지 않음 (장비 미설치)
	i_sIpAddr		: STRING(15);
	i_nPort			: UINT := 502;
	i_nUnitId		: BYTE := 1;
	i_tTimeout		: TIME := T#1S;
END_VAR
VAR_OUTPUT
	q_stState		: ST_TempHumState;		// 읽은 값 (보고 매핑 FB_RptTempHum이 씀)
END_VAR
VAR
	_fbIr			: FB_MBReadInputRegs;
	_awIr			: ARRAY[0..4] OF WORD;	// IR 0..4
	_bReadDue		: BOOL;
	_bReading		: BOOL;
	_bDataOk		: BOOL;					// 한 번이라도 읽음
	_bProbeOk		: BOOL;					// 온도·습도 값이 32767이 아님
END_VAR
VAR CONSTANT
	READ_QTY		: UINT := 5;
	NO_PROBE		: WORD := 16#7FFF;		// 프로브 없음
END_VAR

ACTION A_Map:
_bProbeOk		:= _awIr[1] <> NO_PROBE AND _awIr[2] <> NO_PROBE;
q_stState.fTemp	:= INT_TO_REAL(WORD_TO_INT(_awIr[1])) * 0.01;	// @MAP IR 1 S16 ×0.01 ℃
q_stState.fHum	:= INT_TO_REAL(WORD_TO_INT(_awIr[2])) * 0.01;	// @MAP IR 2 S16 ×0.01 %
_bDataOk := TRUE;
END_ACTION

METHOD M_Cycle
_bReadDue := M_IsReadTime();
IF NOT _bReading THEN
	IF i_bEnable AND i_sIpAddr <> '' AND _bReadDue THEN
		_fbIr(sIPAddr := i_sIpAddr, nTCPPort := i_nPort, nUnitID := i_nUnitId,
			nQuantity := READ_QTY, nMBAddr := 0, cbLength := SIZEOF(_awIr),
			pDestAddr := ADR(_awIr), tTimeout := i_tTimeout, bExecute := TRUE);
		_bReading := TRUE;
	END_IF
ELSE
	_fbIr(bExecute := FALSE);
	IF NOT _fbIr.bBusy THEN
		IF NOT _fbIr.bError AND i_bEnable THEN
			A_Map();
			M_MarkAlive();
		END_IF
		_bReading := FALSE;
	END_IF
END_IF
M_UpdateComm();
q_stState.bValid := Comm AND _bDataOk AND _bProbeOk;
END_METHOD

METHOD M_GetBit : BOOL		// DI 1 값 이상 (통신은 정상인데 프로브 값 무효)
VAR_INPUT
	i_nPoint	: UINT;
END_VAR
IF i_nPoint = 1 THEN
	M_GetBit := Comm AND _bDataOk AND NOT _bProbeOk;
END_IF
END_METHOD

METHOD M_GetValue : ST_Val		// AI 1 온도 ℃, AI 2 습도 %
VAR_INPUT
	i_nPoint	: UINT;
END_VAR
CASE i_nPoint OF
	1:
		M_GetValue.fValue := q_stState.fTemp;
		M_GetValue.bValid := q_stState.bValid;
	2:
		M_GetValue.fValue := q_stState.fHum;
		M_GetValue.bValid := q_stState.bValid;
END_CASE
END_METHOD

METHOD M_SetBit		// 출력 없음
VAR_INPUT
	i_nPoint	: UINT;
	i_bValue	: BOOL;
END_VAR
;
END_METHOD

METHOD M_SetValue		// 출력 없음
VAR_INPUT
	i_nPoint	: UINT;
	i_fValue	: REAL;
END_VAR
;
END_METHOD

PROPERTY Comm : BOOL
GET
Comm := _bComm AND i_bEnable;
END_GET
END_PROPERTY

END_FUNCTION_BLOCK

// ---- 20_Module/Driver/Woonyoung/FB_WoonyoungGfr.TcPOU
FUNCTION_BLOCK FB_WoonyoungGfr EXTENDS FB_DeviceBase IMPLEMENTS I_AuxDevice		// 운영(Woonyoung) WYGF-D08/12/16NC 디지털 지락검출계전기 (Modbus RTU), 읽기 전용
(* ---------------------------------------------------------------
   기반 없음(신규). 맵: 프로토콜 맵 v3\지락검출 계전기.pdf (사용설명서 PAC-00084 REV.5, 제5장). 2026-11-10
   용도: AC 회로 누전(지락) 감시. ZCT 영상변류기 방식이라 배터리 DC 전로 지락은 못 봄 (DC는 IMD)
   통신: EL6022 채널 하나를 ModbusRtuMaster_KL6x22B로 (사용자 2026-11-10). 단자 연결(InData·OutData)은 XAE I/O 화면에서 사람이 함
         장비: RS-485 8N1, 국번 1~32 (공장 출하 OFF → 장비 Serial Setup에서 켜야 응답), 9600/19200/38400 (출하 19200)
   읽기: 읽기 주기마다 Input Register(FC4) 0부터 2 + 회로 수
     @MAP IR 0      U16  시스템 상태 (b8 시험 모드, b4 LPF, b3 고감도 ZCT, b2 자동복귀, b1 부저, b0 50Hz)
     @MAP IR 1      U16  회로별 지락 (b0 = 1회로 … b15 = 16회로, 1 = Fault)
     @MAP IR 2~17   U16  회로 1~16 누설전류, × 0.01 A (예: 0x03E8 = 10 A)
   쓰지 않는 것: FC03 0~31 회로별 감도·동작시간 설정, FC03 32~51 사고 기록, FC05 0 사고 기록 지우기
   점 (I_AuxDevice)
     AI n = 회로 n 누설전류 (A)
     DI n = 회로 n 지락 (n = 1..회로 수), DI 17 = 시험 모드 (장비에서 Circuit Test 중)
   --------------------------------------------------------------- *)
VAR_INPUT
	i_bEnable		: BOOL;					// FALSE면 통신하지 않음 (장비 미설치)
	i_nUnitId		: UINT := 1;			// 장비 국번 (Serial Setup Port No.)
	i_nChannels		: UINT := 8;			// 회로 수: 8 (D08NC), 12 (D12NC), 16 (D16NC)
	i_tTimeout		: TIME := T#1S;			// 응답 기다림
END_VAR
VAR_OUTPUT
	q_wStatus		: WORD;					// IR 0 시스템 상태
	q_wFault		: WORD;					// IR 1 회로별 지락 비트
	q_afCurrent		: ARRAY[1..16] OF REAL;	// 회로별 누설전류 A
	q_bValid		: BOOL;					// 통신 정상이고 한 번 이상 읽음
END_VAR
VAR
	_fbRtu			: ModbusRtuMaster_KL6x22B;
	_awRaw			: ARRAY[0..17] OF WORD;	// IR 0..17
	_bReadDue		: BOOL;
	_bReading		: BOOL;
	_bDataOk		: BOOL;
	_nCh			: UINT;					// 쓰는 회로 수 (8·12·16 중 가까운 범위로 자름)
	_i				: UINT;
END_VAR
VAR CONSTANT
	CH_MAX			: UINT := 16;
	PT_TEST			: UINT := 17;			// DI 17 = 시험 모드
END_VAR

ACTION A_Map:
q_wStatus := _awRaw[0];				// @MAP IR 0
q_wFault := _awRaw[1];				// @MAP IR 1
FOR _i := 1 TO CH_MAX DO
	IF _i <= _nCh THEN
		q_afCurrent[_i] := WORD_TO_REAL(_awRaw[1 + _i]) * 0.01;	// @MAP IR 2~17 U16 ×0.01 A
	ELSE
		q_afCurrent[_i] := 0.0;
	END_IF
END_FOR
_bDataOk := TRUE;
END_ACTION

METHOD M_Cycle
_nCh := LIMIT(1, i_nChannels, CH_MAX);

_bReadDue := M_IsReadTime();
IF NOT _bReading THEN
	IF i_bEnable AND _bReadDue AND i_nUnitId >= 1 AND i_nUnitId <= 247 THEN
		_fbRtu.ReadInputRegs(UnitID := UINT_TO_BYTE(i_nUnitId), Quantity := 2 + _nCh, MBAddr := 0,
			cbLength := SIZEOF(_awRaw), pMemoryAddr := ADR(_awRaw), Timeout := i_tTimeout, Execute := TRUE);
		_bReading := TRUE;
	END_IF
ELSE
	_fbRtu.ReadInputRegs(Execute := FALSE);	// 시작한 읽기는 끝까지 부름
	IF NOT _fbRtu.BUSY THEN
		IF NOT _fbRtu.Error AND i_bEnable THEN
			A_Map();
			M_MarkAlive();
		END_IF
		_bReading := FALSE;
	END_IF
END_IF
M_UpdateComm();
q_bValid := Comm AND _bDataOk;
END_METHOD

METHOD M_GetBit : BOOL		// DI n = 회로 n 지락, DI 17 = 시험 모드. 통신 이상이면 FALSE (규칙 FB_RuleBit은 Comm으로 따로 판단)
VAR_INPUT
	i_nPoint	: UINT;
END_VAR
IF q_bValid THEN
	IF i_nPoint >= 1 AND i_nPoint <= _nCh THEN
		M_GetBit := (q_wFault AND SHL(WORD#1, i_nPoint - 1)) <> 0;
	ELSIF i_nPoint = PT_TEST THEN
		M_GetBit := q_wStatus.8;
	END_IF
END_IF
END_METHOD

METHOD M_GetValue : ST_Val		// AI n = 회로 n 누설전류 (A)
VAR_INPUT
	i_nPoint	: UINT;
END_VAR
IF i_nPoint >= 1 AND i_nPoint <= _nCh THEN
	M_GetValue.fValue := q_afCurrent[i_nPoint];
	M_GetValue.bValid := q_bValid;
END_IF
END_METHOD

METHOD M_SetBit		// 출력 없음
VAR_INPUT
	i_nPoint	: UINT;
	i_bValue	: BOOL;
END_VAR
;
END_METHOD

METHOD M_SetValue		// 출력 없음
VAR_INPUT
	i_nPoint	: UINT;
	i_fValue	: REAL;
END_VAR
;
END_METHOD

PROPERTY Comm : BOOL
GET
Comm := _bComm AND i_bEnable;
END_GET
END_PROPERTY

END_FUNCTION_BLOCK

// ---- 20_Module/Driver/Gasdna/FB_GasdnaAsd57.TcPOU
FUNCTION_BLOCK FB_GasdnaAsd57 EXTENDS FB_DeviceBase IMPLEMENTS I_AuxDevice		// 가스디엔에이 ASD-57 열연복합 감지기 (Modbus RTU), 읽기 전용
(* ---------------------------------------------------------------
   기반 없음(신규). 맵: 프로토콜 맵 v3\ASD-5x(모드 버스 프로토콜)_ver1.1(22_0922).pdf, 결선: ASD-57_매뉴얼.pdf. 2026-11-10
   통신: EL6022 채널 하나를 ModbusRtuMaster_KL6x22B로. 단자 연결(InData·OutData)은 XAE I/O 화면에서 사람이 함
         장비: RS-485 9600 bps 고정, 8N1, 국번 1~126 (출하 1). 흰 TX+, 파랑 TX-
         속도가 9600 고정이라 다른 속도 장비(지락계전기 출하 19200)와 한 채널에 묶지 않음
         응답 뒤 10 ms 이상 지나 다음 요청 (읽기 주기 1 s라 맞음)
   읽기: 읽기 주기마다 Holding Register(FC3) 0부터 9칸
     @MAP HR 0 (40001) U16  1 Color 연기 농도 0~1000, ×0.1 %
     @MAP HR 1 (40002) U16  2 Color 연기 농도 0~1000, ×0.01 (맵 표기 x.xx, 단위 표기 없음)
     @MAP HR 2 (40003) U16  온도 0~1000, ×0.1 ℃ (ASD-57 전용)
     @MAP HR 3 (40004) U16  알람 상태: 0 없음, 1 연기 (1·2 Color 모두 알람값 초과), 2 온도 (ASD-57 전용)
     @MAP HR 4 (40005) U16  1 Color 연기 알람값 (출하 80)
     @MAP HR 5 (40006) U16  2 Color 연기 알람값 (출하 170)
     @MAP HR 6 (40007) U16  온도 알람값 ×0.1 ℃ (출하 700 = 70.0 ℃)
     @MAP HR 7 (40008) U16  딜레이 ×10 ms (최대 1000 = 10 s)
     @MAP HR 8 (40009) U16  통신 국번
   쓰지 않는 것: FC6 HR 4~8 설정 바꾸기, HR 50 ZERO 교정(1234). 설정은 장비 출하값 그대로 (바꾸려면 사용자 결정)
   알람 상태 3(연기 + 온도)은 맵에 없음 → 비트로 봄 (b0 연기, b1 온도)
   점 (I_AuxDevice)
     AI 1 = 1 Color 연기 %, AI 2 = 2 Color 연기, AI 3 = 온도 ℃
     DI 1 = 연기 알람, DI 2 = 온도 알람
   --------------------------------------------------------------- *)
VAR_INPUT
	i_bEnable		: BOOL;					// FALSE면 통신하지 않음 (장비 미설치)
	i_nUnitId		: UINT := 1;			// 장비 국번 (HR 8)
	i_tTimeout		: TIME := T#1S;			// 응답 기다림
END_VAR
VAR_OUTPUT
	q_fSmoke1		: REAL;					// 1 Color 연기 농도 %
	q_fSmoke2		: REAL;					// 2 Color 연기 농도
	q_fTemp			: REAL;					// 온도 ℃
	q_wAlarm		: WORD;					// HR 3 알람 상태 원시값
	q_bSmokeAlarm	: BOOL;					// 연기 알람
	q_bTempAlarm	: BOOL;					// 온도 알람
	q_anSet			: ARRAY[4..8] OF UINT;	// HR 4~8 설정값 원시값 (알람값, 딜레이, 국번)
	q_bValid		: BOOL;					// 통신 정상이고 한 번 이상 읽음
END_VAR
VAR
	_fbRtu			: ModbusRtuMaster_KL6x22B;
	_awRaw			: ARRAY[0..8] OF WORD;	// HR 0..8
	_bReadDue		: BOOL;
	_bReading		: BOOL;
	_bDataOk		: BOOL;
	_i				: UINT;
END_VAR
VAR CONSTANT
	READ_QTY		: UINT := 9;
END_VAR

ACTION A_Map:
q_fSmoke1 := WORD_TO_REAL(_awRaw[0]) * 0.1;		// @MAP HR 0 ×0.1 %
q_fSmoke2 := WORD_TO_REAL(_awRaw[1]) * 0.01;	// @MAP HR 1 ×0.01
q_fTemp := WORD_TO_REAL(_awRaw[2]) * 0.1;		// @MAP HR 2 ×0.1 ℃
q_wAlarm := _awRaw[3];							// @MAP HR 3
q_bSmokeAlarm := q_wAlarm.0;
q_bTempAlarm := q_wAlarm.1;
FOR _i := 4 TO 8 DO
	q_anSet[_i] := WORD_TO_UINT(_awRaw[_i]);	// @MAP HR 4~8
END_FOR
_bDataOk := TRUE;
END_ACTION

METHOD M_Cycle
_bReadDue := M_IsReadTime();
IF NOT _bReading THEN
	IF i_bEnable AND _bReadDue AND i_nUnitId >= 1 AND i_nUnitId <= 126 THEN
		_fbRtu.ReadRegs(UnitID := UINT_TO_BYTE(i_nUnitId), Quantity := READ_QTY, MBAddr := 0,
			cbLength := SIZEOF(_awRaw), pMemoryAddr := ADR(_awRaw), Timeout := i_tTimeout, Execute := TRUE);
		_bReading := TRUE;
	END_IF
ELSE
	_fbRtu.ReadRegs(Execute := FALSE);	// 시작한 읽기는 끝까지 부름
	IF NOT _fbRtu.BUSY THEN
		IF NOT _fbRtu.Error AND i_bEnable THEN
			A_Map();
			M_MarkAlive();
		END_IF
		_bReading := FALSE;
	END_IF
END_IF
M_UpdateComm();
q_bValid := Comm AND _bDataOk;
END_METHOD

METHOD M_GetBit : BOOL		// DI 1 연기 알람, DI 2 온도 알람. 통신 이상이면 FALSE (규칙 FB_RuleBit은 Comm으로 따로 판단)
VAR_INPUT
	i_nPoint	: UINT;
END_VAR
IF q_bValid THEN
	CASE i_nPoint OF
		1: M_GetBit := q_bSmokeAlarm;
		2: M_GetBit := q_bTempAlarm;
	END_CASE
END_IF
END_METHOD

METHOD M_GetValue : ST_Val		// AI 1 연기1 %, AI 2 연기2, AI 3 온도 ℃
VAR_INPUT
	i_nPoint	: UINT;
END_VAR
CASE i_nPoint OF
	1: M_GetValue.fValue := q_fSmoke1;
	2: M_GetValue.fValue := q_fSmoke2;
	3: M_GetValue.fValue := q_fTemp;
ELSE
	RETURN;
END_CASE
M_GetValue.bValid := q_bValid;
END_METHOD

METHOD M_SetBit		// 출력 없음
VAR_INPUT
	i_nPoint	: UINT;
	i_bValue	: BOOL;
END_VAR
;
END_METHOD

METHOD M_SetValue		// 출력 없음
VAR_INPUT
	i_nPoint	: UINT;
	i_fValue	: REAL;
END_VAR
;
END_METHOD

PROPERTY Comm : BOOL
GET
Comm := _bComm AND i_bEnable;
END_GET
END_PROPERTY

END_FUNCTION_BLOCK

// ---- 20_Module/Virtual/FB_SrcTest.TcPOU
FUNCTION_BLOCK FB_SrcTest EXTENDS FB_SourceBase		// 시험 지령원: 온라인으로 값을 써서 시험
VAR_INPUT
	i_ePcsReq			: E_PcsCmd;		// PCS 요청. 쓰면 1스캔 요청으로 나가고 None으로 돌아감
	i_nPcsUnit			: UINT;			// 0 = 그룹 전체, n = 유닛 n
	i_eBatReq			: E_BatCmd;		// 배터리 요청 (Close / Open). 쓰면 1스캔 요청으로 나가고 None으로 돌아감
	i_nBatGroup			: UINT;			// 0 = 전체, n = 배터리 그룹 n
	i_bPSetActive		: BOOL;
	i_fPSet				: REAL;			// kW, 접속점 기준 (방전 +)
	i_bQSetActive		: BOOL;
	i_fQSet				: REAL;			// kvar, 접속점 기준 (공급 +)
	i_bPLimActive		: BOOL;			// 지령원 P 제한 시험
	i_fPMax				: REAL;			// kW
	i_fPMin				: REAL;
	i_bQLimActive		: BOOL;			// 지령원 Q 제한 시험
	i_fQMax				: REAL;			// kvar
	i_fQMin				: REAL;
	(* 유닛별 값 시험 (유닛 하나) *)
	i_nUnit				: UINT;			// 0 = 안 씀
	i_bUnitPSetActive	: BOOL;
	i_fUnitPSet			: REAL;			// kW, 유닛 출력
	i_bSend				: BOOL;			// 같은 값을 다시 보낼 때 TRUE (값을 바꾸면 자동으로 새 지령)
END_VAR

METHOD M_UpdateOutput : BOOL
VAR
	u		: UINT;
	stOld	: ST_SourceOutput;
END_VAR
stOld := _stOut;

_stOut.bPSetActive	:= i_bPSetActive;
_stOut.fPSet		:= i_fPSet;
_stOut.bQSetActive	:= i_bQSetActive;
_stOut.fQSet		:= i_fQSet;
_stOut.bPLimActive	:= i_bPLimActive;
_stOut.fPMax		:= i_fPMax;
_stOut.fPMin		:= i_fPMin;
_stOut.bQLimActive	:= i_bQLimActive;
_stOut.fQMax		:= i_fQMax;
_stOut.fQMin		:= i_fQMin;
IF i_ePcsReq <> E_PcsCmd.None THEN
	_stOut.stPcsReq.eCmd	:= i_ePcsReq;
	_stOut.stPcsReq.nUnit	:= i_nPcsUnit;
	i_ePcsReq				:= E_PcsCmd.None;
END_IF
IF i_eBatReq <> E_BatCmd.None THEN
	_stOut.stBatReq.eCmd		:= i_eBatReq;
	_stOut.stBatReq.nBatGroup	:= i_nBatGroup;
	i_eBatReq					:= E_BatCmd.None;
END_IF

